(* IEC 61131-3 sources: daoli-st-library/DL_Motion (part 2) *)

(* ---- FB_DL_ResolverEncoderRedundSwitch.st ---- *)
(*
    FB_DL_ResolverEncoderRedundSwitch —— 旋变 + 增量编码器双通道角反馈冗余判定与无扰切换
    ------------------------------------------------------------------
    组件名    : FB_DL_ResolverEncoderRedundSwitch
    分类      : DL_Motion / Feedback Redundancy（反馈冗余切换）
    一句话功能: 双通道角反馈偏差超限时判定哪一路可信并无扰切到单通道运行，
                切换过程中输出角度受变率限制，绝不产生位置跳变。
    复杂度    : C4
    版本      : v1.0.0
    开源溯源  : 无（clean-room 自研，未借鉴任何开源实现）
    平台      : 纯 IEC 61131-3（TON / R_TRIG / ABS / REAL_TO_INT / INT_TO_REAL 标准转换），
                目标编译器 RuSTy 1.0.8，兼容 CODESYS 3.5 / TwinCAT 3 / 汇川 InoProShop /
                Machine Expert；无 PROPERTY、无 VLA、无 FOR..DOWNTO、无 AS 类方言
    ------------------------------------------------------------------
    功能说明  : ① 角差按 360° 环形折算：先各自折到 [0,360)，再
                   d := ABS(fAngleA − fAngleB)；IF d > 180 THEN d := 360 − d（结果域 [0,180]）；
                ② 双通道都有效且角差在容差内 → 融合输出（两路短弧中点），并每拍刷新
                   「融合参照角」_fRefDeg，供后续判定「哪一路可信」时作参照；
                ③ 角差超容差且持续 tFaultPersistMs（TON 无条件刷新）→ 判 SUSPECT；
                   任一路 bXValid = FALSE（或该路角度非有限）→ 直接判该路失效并切单通道；
                ④ 判定「哪一路可信」：以「最近一次双通道合格时的融合参照角」为准，
                   取与参照偏离较小者（相等时稳定优先取旋变 A）；无参照 → LOST，不猜；
                ⑤ 切换时 fAngleOut 按 fMaxSlewDegPerSec 限变率跟随目标角：环形带符号差值
                   先钳到 ±每拍步长再累加，故任何切换都不产生跳变；
                ⑥ 输出通道码 nActiveChannel：0 = 融合、1 = 旋变 A、2 = 编码器 B、-1 = 无。
    量纲链    : fAngleADeg [°] − fAngleBDeg [°] → 角差 [°]（经 360° 折算，域 [0,180]）；
                _fDevRatio = _fDevDeg [°] ÷ _fTolGuard [°] → 无因次 [-]（故与 1.0 直比判超限）；
                fMaxSlewDegPerSec [°/s] × DL_RE_SAMPLE_S [s] → 每拍最大角增量 [°]；
                _fDelta [°] 钳到 ±步长 [°] 后加到 _fOut [°] 再折回 [0,360) → fAngleOut [°]。
                全程无「角度与时间相加」「比例与角度相加」，量纲链逐段闭合。
    代理假设  : （R95 三句声明）① 代理值 = 常量 DL_RE_SAMPLE_S = 0.004 s，代表本 FB 所在
                任务的标称扫描周期；② 覆盖范围 = 2 ms ~ 10 ms 的周期任务（最坏 ±60% 误差只
                影响切换变率的平滑度，不改变安全判据的判定结果）；③ 覆盖不到的区间
                （< 1 ms 高速任务、事件任务、扫描周期抖动超 10 ms）由驱动层位置环限幅与伺服
                自身加速度限制负责，本件限变率只作二级防线。
    交付门槛  : 本件使用 REAL_TO_INT / INT_TO_REAL 标准转换做角度折圈，须在 CODESYS /
                TwinCAT / InoProShop 三平台各编译验证一次（R64）。
    状态机    : eInit(0) --双路有效且角差在容差内--> eDualOk(10)
                eInit --双路有效但角差超限--> eSuspect(20)；--仅一路有效--> eSingleA(30)/eSingleB(40)
                eDualOk --角差超容差持续 tFaultPersistMs 到（tonDev.Q）--> eSuspect
                eDualOk/eSuspect --A 失效--> eSingleB；--B 失效--> eSingleA
                eSuspect --有参照且可判--> eSingleA/eSingleB；--无参照或双路皆失效--> eLost(90)
                eSingleA/eSingleB --对侧恢复且一致计时到（tonAgree.Q）--> eDualOk
                eSingleA --A 失效--> eLost；eSingleB --B 失效--> eLost
                eLost --双路恢复且一致计时到（tonAgree.Q）--> eDualOk；
                eLost --单路恢复且确认计时到（tonSingle.Q）--> eSingleA/eSingleB（先进单通道，不直接回双通道）
                解除路径自证：tonSingle 的 IN 为「恰好一路可用」，故 eLost 的单路恢复边恒可达；
                若两路长期不一致且从未建立参照，eLost 按设计保持（不猜），bReset 重建参照后再裁决
    失能语义  : bEnable = FALSE 时 eState := eInit、nActiveChannel := -1、bLost := FALSE，
                fAngleOut 冻结保持末值（不跳变、不清零）；恢复使能后按变率追随新目标角。
                取「冻结保持」而非「降级清零」：角度是位置事实量，清零等于伪造位置（R191）。
    复位作用域: bReset 上升沿①清 _fRefDeg 与 _bRefValid（参照作废，须重建双通道合格）；
                ②清 _bCfgBad 与各成因位；③迁相回 eInit；④不清 _fOut（角度不得因复位跳变）。
    防御口径  : NaN 用自反 f<>f；±Inf 用 (f−f)<>(f−f)；另设幅值域闸 ABS(f) > 1.0E30。
                折圈除法的除子为常量 360.0（无零风险），但实数转整数前先做幅值域钳制，防
                REAL_TO_INT 溢出翻转（R151）；容差比值除法先以 DL_RE_TOL_FLOOR 两级兜底除子。
    规格补充  : 派单引脚表未含变率限制引脚，但设计要求「输出必须限变率」，故补充输入
                fMaxSlewDegPerSec（默认 3600 °/s，即 10 圈每秒）。派单写作 iActiveChannel（INT）；
                本库命名规范 1.2 规定有符号整数前缀为 n、i 专用于接口引用，故落为
                nActiveChannel，语义与码值一字不减。另按 R190 归因唯一补充 bCfgErr / bDataErr
                两个诊断位，使「组态非法」与「通道数据非有限」两条成因各自可观测。
    码位说明  : 本件按零码位范式交付，不分配 16# 事件码；失效成因（A 失效 / B 失效 /
                双路同时失效 / 无参照 / 当前通道失效 / 组态非法）各有独立内部成员，
                经 eState 与 bLost 观测，不共用同一枚举成员归因（R190）。
    修订记录  : 2026-11-24 v1.0.0 首次入库（R87 批 · #2）
*)
TYPE E_DL_ResEncState :
(
    eInit    := 0,    // 初始化或未投运：输出冻结，不判角差 | init or disabled, output frozen, no judging
    eDualOk  := 10,   // 双通道合格：融合输出，刷新融合参照角 | dual channels healthy, fused output, reference refreshed
    eSuspect := 20,   // 疑似：角差持续超容差，正在判定可信通道 | suspect, deviation persisted, arbitrating the trusted channel
    eSingleA := 30,   // 单通道 A：仅旋变通道参与输出 | single channel A, resolver only
    eSingleB := 40,   // 单通道 B：仅编码器通道参与输出 | single channel B, encoder only
    eLost    := 90    // 失效：无可信通道或无参照可判，输出冻结 | lost, no trusted channel or no reference
);
END_TYPE

FUNCTION_BLOCK FB_DL_ResolverEncoderRedundSwitch
VAR_INPUT
    bEnable            : BOOL;                    // 使能电平，TRUE = 允许切换判定 | enable level, TRUE = arbitration active
    bReset             : BOOL;                    // 复位请求，上升沿生效 | reset request, rising-edge active
    fAngleADeg         : REAL;                    // 旋变通道角度 [°]，任意圈数，内部折到 0..360 | resolver angle [deg]
    fAngleBDeg         : REAL;                    // 增量编码器角度 [°]，任意圈数，内部折到 0..360 | encoder angle [deg]
    fTolDeg            : REAL := 0.5;             // 双通道允许角差 [°]，须为正 | allowed channel deviation [deg]
    tFaultPersistMs    : TIME := T#100MS;         // 超限与恢复一致的持续确认时长 [ms] | persistence time [ms]
    bAValid            : BOOL;                    // 旋变通道有效位，驱动侧给出 | resolver channel validity from the drive
    bBValid            : BOOL;                    // 编码器通道有效位，驱动侧给出 | encoder channel validity from the drive
    fMaxSlewDegPerSec  : REAL := 3600.0;          // 输出角度最大变率 [°/s]，须为正 | max output slew rate [deg/s]
END_VAR
VAR_OUTPUT
    eState             : E_DL_ResEncState;        // 主状态，供 HMI 与联锁使用 | main state for HMI and interlocks
    fAngleOut          : REAL;                    // 参与位置环的输出角度 [°]，域 [0,360) 且限变率 | output angle [deg]
    fDeviationDeg      : REAL;                    // 本拍环形角差 [°]，域 [0,180] | circular deviation this scan [deg]
    nActiveChannel     : INT;                     // 通道码：0 融合 / 1 旋变 A / 2 编码器 B / -1 无 | channel code
    bSwitchEvent       : BOOL;                    // 通道切换事件位，单拍 | channel switch event, single scan
    bLost              : BOOL;                    // 失效汇总位，eLost 相为 TRUE | lost aggregate, TRUE in the eLost phase
    bCfgErr            : BOOL;                    // 组态非法诊断位（归因唯一，R190）| bad-configuration flag, unique attribution
    bDataErr           : BOOL;                    // 数据非有限诊断位（归因唯一，R190）| non-finite data flag, unique attribution
END_VAR
VAR
    rtReset            : R_TRIG;                  // 复位上升沿实例，每拍无条件刷新 | reset rising-edge instance
    tonDev             : TON;                     // 角差超限持续确认计时，每拍无条件刷新 | deviation persistence timer
    tonAgree           : TON;                     // 双通道一致确认计时，每拍无条件刷新 | agreement persistence timer
    tonSingle          : TON;                     // 单通道恢复确认计时，每拍无条件刷新 | single-channel recovery timer
    _eState            : E_DL_ResEncState := E_DL_ResEncState.eInit; // 状态机内部当前态 | internal current state
    _bInit             : BOOL := TRUE;            // 首扫初始化标志，含参照与输出保持槽状态 | first-scan init flag
    _bResetLatch       : BOOL := FALSE;           // 复位沿锁存量，本拍末清除 | reset-edge latch, cleared at scan end
    _bCfgBad           : BOOL := FALSE;           // 组态非法标志 | bad configuration flag
    _bAOk              : BOOL := FALSE;           // 旋变通道可用（有效位且角度有限）| resolver channel usable
    _bBOk              : BOOL := FALSE;           // 编码器通道可用（有效位且角度有限）| encoder channel usable
    _bLostBoth         : BOOL := FALSE;           // 双路同时失效成因位（归因唯一）| both channels lost
    _bNoRef            : BOOL := FALSE;           // 无融合参照成因位（归因唯一）| no reference available
    _bChLost           : BOOL := FALSE;           // 当前单通道失效成因位（归因唯一）| the active single channel was lost
    _fOut              : REAL := 0.0;             // 输出角度保持槽 [°]，域 [0,360) | output angle holder [deg]
    _fRefDeg           : REAL := 0.0;             // 融合参照角 [°]，仅在双通道合格时刷新 | fused reference angle [deg]
    _bRefValid         : BOOL := FALSE;           // 融合参照角可用标志 | fused reference valid flag
    _fDevDeg           : REAL := 0.0;             // 本拍环形角差 [°] | circular deviation this scan [deg]
    _fDevRatio         : REAL := 0.0;             // 角差与容差之比 [-]，判超限用 | deviation to tolerance ratio
    _fTolGuard         : REAL := 0.0;             // 带下限兜底的容差 [°]，作除法除子 | tolerance with floor, used as divisor
    _fSlewStep         : REAL := 0.0;             // 每拍最大角增量 [°] | max angle increment per scan [deg]
    _fDelta            : REAL := 0.0;             // 本拍待施加带符号角增量 [°]（已钳位）| clamped angle increment [deg]
    _fTarget           : REAL := 0.0;             // 本拍目标角 [°] | target angle this scan [deg]
    _fFuse             : REAL := 0.0;             // 本拍融合角 [°] | fused angle this scan [deg]
    _fDevA             : REAL := 0.0;             // A 相对参照的偏离 [°] | A deviation from the reference [deg]
    _fDevB             : REAL := 0.0;             // B 相对参照的偏离 [°] | B deviation from the reference [deg]
    _nCh               : INT := -1;               // 本拍通道码 | channel code this scan
    _nChPrev           : INT := -1;               // 上一拍通道码，供切换事件差分 | previous channel code for the switch event
    nFoldIdx           : INT := 0;                // 折圈方法内残余修正循环下标 | residue loop index inside the folding method
END_VAR
VAR CONSTANT
    DL_RE_EPS          : REAL := 1.0E-6;          // 浮点判零容差 [°] | float zero tolerance [deg]
    DL_RE_TOL_FLOOR    : REAL := 1.0E-4;          // 容差参数下限兜底 [°] | tolerance floor [deg]
    DL_RE_MAG_MAX      : REAL := 1.0E30;          // 有限幅值域闸上限（角度与变率）[°] | magnitude domain bound [deg]
    DL_RE_FOLD_MAX     : REAL := 1.0E6;           // 折圈前的角度幅值域上限 [°]，实数转整数前钳制 | fold domain bound [deg]
    DL_RE_SAMPLE_S     : REAL := 0.004;           // 代理扫描周期 [s]，见头注释代理假设三句 | proxy sample period [s]
    DL_RE_DEG_FULL     : REAL := 360.0;           // 整圈角度 [°] | full turn [deg]
    DL_RE_DEG_HALF     : REAL := 180.0;           // 半圈角度 [°] | half turn [deg]
    DL_RE_FUSE_W       : REAL := 0.5;             // 融合权重，两路等权且权值和为 1 [-] | fusion weight, sums to one
    DL_RE_CH_FUSE      : INT := 0;                // 通道码：融合 | channel code, fused
    DL_RE_CH_A         : INT := 1;                // 通道码：旋变 A | channel code, resolver A
    DL_RE_CH_B         : INT := 2;                // 通道码：编码器 B | channel code, encoder B
    DL_RE_CH_NONE      : INT := -1;               // 通道码：无 | channel code, none
    DL_RE_FOLD_ITER    : INT := 8;                // 折圈残余修正最大迭代次数（防死循环计数器）| fold iteration guard
END_VAR

METHOD FoldAngleDeg : REAL
(*
    角度折圈：把任意圈数角度折到 [0,360)。先按幅值域钳制再转整数，防 REAL_TO_INT 溢出翻转。
    Angle folding into [0,360): the magnitude is bounded before the real-to-integer conversion.
*)
VAR_INPUT
    fIn : REAL;                                   // 待折圈角度 [°] | angle to fold [deg]
END_VAR
VAR
    nTurn : INT;                                  // 整圈数，截断取整后按符号修正 [-] | whole turns after truncation
END_VAR
IF (fIn <> fIn) OR ((fIn - fIn) <> (fIn - fIn)) THEN
    FoldAngleDeg := 0.0;                          // NaN 或 ±Inf：返回哨兵零点，由调用方闸门拦截 | non-finite input returns the sentinel zero
    RETURN;
END_IF
IF (fIn > DL_RE_FOLD_MAX) OR (fIn < (0.0 - DL_RE_FOLD_MAX)) THEN
    FoldAngleDeg := 0.0;                          // 超折圈域：返回哨兵零点不猜，域外由上游闸门负责 | out of fold domain, return the sentinel
    RETURN;
END_IF
nTurn := REAL_TO_INT(fIn / DL_RE_DEG_FULL);       // 圈数 [-] = [°] ÷ 常量 360.0（除子为常量，无除零风险）| turns, constant divisor
FoldAngleDeg := fIn - INT_TO_REAL(nTurn) * DL_RE_DEG_FULL; // 折圈结果 [°] = [°] − [-] × [°] | folded angle [deg]
FOR nFoldIdx := 1 TO DL_RE_FOLD_ITER DO
    IF FoldAngleDeg < 0.0 THEN
        FoldAngleDeg := FoldAngleDeg + DL_RE_DEG_FULL; // 负角补整圈 [°] | add one turn for negative angles
    END_IF
END_FOR
IF FoldAngleDeg >= DL_RE_DEG_FULL THEN
    FoldAngleDeg := 0.0;                          // 折圈后仍越上界（数值极值退化）：返回哨兵零点 | degenerate result returns the sentinel
END_IF
END_METHOD

METHOD FoldDeviationDeg : REAL
(*
    环形角差幅值：d := ABS(A − B)；IF d > 180 THEN d := 360 − d，结果域 [0,180]（派单指定口径）。
    Circular deviation magnitude, exactly the formula requested by the dispatch.
*)
VAR_INPUT
    fAngleA : REAL;                               // A 通道角度 [°] | channel A angle [deg]
    fAngleB : REAL;                               // B 通道角度 [°] | channel B angle [deg]
END_VAR
VAR
    fD : REAL;                                    // 角差中间量 [°] | deviation intermediate [deg]
END_VAR
fD := ABS(FoldAngleDeg(fAngleA) - FoldAngleDeg(fAngleB)); // 折圈后作差取绝对值 [°] | absolute difference of folded angles
IF fD > DL_RE_DEG_HALF THEN
    fD := DL_RE_DEG_FULL - fD;                    // 折到短弧侧 [°]，与派单口径一致 | fold onto the short arc [deg]
END_IF
FoldDeviationDeg := fD;
END_METHOD

METHOD FoldSignedDiff : REAL
(*
    环形带符号差：返回 A − B 折到 (-180, 180]，用于融合与限变率增量计算。
    Signed circular difference folded into (-180, 180], used by fusion and by the slew limiter.
*)
VAR_INPUT
    fAngleA : REAL;                               // 被减角度 [°] | minuend angle [deg]
    fAngleB : REAL;                               // 减数角度 [°] | subtrahend angle [deg]
END_VAR
VAR
    fD : REAL;                                    // 带符号角差中间量 [°] | signed difference intermediate [deg]
END_VAR
fD := FoldAngleDeg(fAngleA) - FoldAngleDeg(fAngleB); // 折圈后作差 [°] | difference of folded angles [deg]
IF fD > DL_RE_DEG_HALF THEN
    fD := fD - DL_RE_DEG_FULL;                    // 折到负侧 [°] | fold into the negative side [deg]
END_IF
IF fD <= (0.0 - DL_RE_DEG_HALF) THEN
    fD := fD + DL_RE_DEG_FULL;                    // 折到正侧 [°] | fold into the positive side [deg]
END_IF
FoldSignedDiff := fD;
END_METHOD

// 段 1｜输出安全侧预置与首扫初始化（含参照与保持槽状态，故必须有 _bInit，R310）
// segment 1, safe-value presets and first-scan initialisation; the reference holder requires _bInit
nActiveChannel := DL_RE_CH_NONE;                   // 预置通道码「无」| preset channel code to none
bLost := FALSE;                                    // 预置未失效 | preset not lost
bSwitchEvent := FALSE;                             // 预置无切换事件 | preset no switch event
_fDevDeg := 0.0;                                   // 预置角差 0 [°] | preset zero deviation [deg]
_fDevRatio := 0.0;                                 // 预置角差比 0 [-] | preset zero ratio
_bCfgBad := FALSE;                                 // 预置组态合法 | preset legal configuration
_bLostBoth := FALSE;                               // 预置双路未同时失效 | preset both channels not lost
_bNoRef := FALSE;                                  // 预置参照缺失未置位 | preset reference-missing flag clear
_bChLost := FALSE;                                 // 预置当前通道未失效 | preset active-channel-lost flag clear
_nCh := DL_RE_CH_NONE;                             // 预置本拍通道码「无」| preset the channel code to none
IF _bInit THEN
    _bInit := FALSE;                               // 首扫只执行一次 | runs once on the first scan
    _eState := E_DL_ResEncState.eInit;             // 首扫状态回初相 | initialise the state
    _bRefValid := FALSE;                           // 参照角作废，须重建 | invalidate the reference
    IF (fAngleADeg <> fAngleADeg) OR ((fAngleADeg - fAngleADeg) <> (fAngleADeg - fAngleADeg)) THEN
        _fOut := 0.0;                              // 首扫角度非有限：保持槽取哨兵零点，等闸门置失效 | non-finite first angle
    ELSE
        _fOut := FoldAngleDeg(fAngleADeg);         // 首扫以旋变角为输出起点 [°]，避免首拍从 0 跳变 | start from the resolver angle
    END_IF
    _nChPrev := DL_RE_CH_NONE;                     // 首扫通道快照为「无」| first-scan channel snapshot
END_IF

// 段 2｜通道可用性判定：有效位 + NaN 自反 + Inf 自减 + 幅值域，逐个浮点入参枚举（R4 / R151 / R272）
// segment 2, channel usability: validity bit plus NaN self-reflexive, Inf self-subtraction and the magnitude bound
_bAOk := bAValid;
IF (fAngleADeg <> fAngleADeg) OR ((fAngleADeg - fAngleADeg) <> (fAngleADeg - fAngleADeg)) THEN
    _bAOk := FALSE;                                // 旋变角 NaN 或 ±Inf：判该路失效 | NaN or infinity, the channel is unusable
END_IF
IF ABS(fAngleADeg) > DL_RE_MAG_MAX THEN
    _bAOk := FALSE;                                // 旋变角超幅值域：判该路失效 | beyond the magnitude domain, unusable
END_IF
_bBOk := bBValid;
IF (fAngleBDeg <> fAngleBDeg) OR ((fAngleBDeg - fAngleBDeg) <> (fAngleBDeg - fAngleBDeg)) THEN
    _bBOk := FALSE;                                // 编码器角 NaN 或 ±Inf：判该路失效 | NaN or infinity, the channel is unusable
END_IF
IF ABS(fAngleBDeg) > DL_RE_MAG_MAX THEN
    _bBOk := FALSE;                                // 编码器角超幅值域：判该路失效 | beyond the magnitude domain, unusable
END_IF

// 段 3｜容差两级兜底与组态闸（容差作除子，必须先兜底再除；变率须为正且有限）
// segment 3, two-stage tolerance fallback and configuration gate; the tolerance is a divisor, floor it first
_fTolGuard := fTolDeg;                             // 取配置容差 [°] | take the configured tolerance [deg]
IF (fTolDeg <> fTolDeg) OR ((fTolDeg - fTolDeg) <> (fTolDeg - fTolDeg)) THEN
    _fTolGuard := DL_RE_TOL_FLOOR;                 // 容差非有限：一级回默认下限 [°] | non-finite tolerance falls back to the floor
END_IF
IF _fTolGuard < DL_RE_TOL_FLOOR THEN
    _fTolGuard := DL_RE_TOL_FLOOR;                 // 容差过小或为负：二级按有效域钳定 [°] | too small or negative, clamp to the floor
END_IF
IF (fMaxSlewDegPerSec <> fMaxSlewDegPerSec) OR ((fMaxSlewDegPerSec - fMaxSlewDegPerSec) <> (fMaxSlewDegPerSec - fMaxSlewDegPerSec)) THEN
    _bCfgBad := TRUE;                              // 变率非有限：组态非法 | non-finite slew rate, illegal configuration
END_IF
IF fMaxSlewDegPerSec <= DL_RE_EPS THEN
    _bCfgBad := TRUE;                              // 变率非正：组态非法（无变率限制即失去无扰切换保障）| non-positive slew rate
END_IF
IF ABS(fMaxSlewDegPerSec) > DL_RE_MAG_MAX THEN
    _bCfgBad := TRUE;                              // 变率超幅值域：组态非法 | slew rate beyond the magnitude domain
END_IF
IF tFaultPersistMs < T#0S THEN
    _bCfgBad := TRUE;                              // 持续确认时长为负：组态非法 | negative persistence time, illegal configuration
END_IF

// 段 4｜本拍角差与角差比（双路都可用才计算，否则记 0 且不参与判据）
// segment 4, deviation and deviation ratio this scan; computed only when both channels are usable
IF _bAOk AND _bBOk THEN
    _fDevDeg := FoldDeviationDeg(fAngleADeg, fAngleBDeg); // 环形角差 [°] | circular deviation [deg]
    _fDevRatio := _fDevDeg / _fTolGuard;           // 角差比 [-] = [°] ÷ [°]，_fTolGuard 已两级兜底非零 | guarded division
ELSE
    _fDevDeg := 0.0;                               // 单路或双路失效：角差无意义记 0 [°] | deviation meaningless here
    _fDevRatio := 0.0;                             // 单路或双路失效：角差比记 0 [-] | ratio meaningless here
END_IF

// 段 5｜定时器与沿实例无条件周期刷新（R7：严禁放入 IF / CASE 分支内部），入参为本拍已算量
// segment 5, timers and edge instances refreshed unconditionally, fed with values already computed this scan
rtReset(CLK := bReset);
tonDev(IN := bEnable AND _bAOk AND _bBOk AND (_fDevRatio > 1.0), PT := tFaultPersistMs);
tonAgree(IN := bEnable AND _bAOk AND _bBOk AND (_fDevRatio <= 1.0), PT := tFaultPersistMs);
tonSingle(IN := bEnable AND (_bAOk OR _bBOk) AND (NOT (_bAOk AND _bBOk)), PT := tFaultPersistMs);
IF rtReset.Q THEN
    _bResetLatch := TRUE;                          // 复位沿存锁存量，段 6 统一消费 | store the reset edge, consumed in segment 6
END_IF

// 段 6｜复位沿处理（先复位后判据，保证本拍新事件不被抹除，R275）
// segment 6, reset edge handling; reset runs before the criteria so same-scan events survive
IF _bResetLatch THEN
    _bRefValid := FALSE;                           // 参照作废，须重新建立双通道合格 | invalidate the reference
    _fRefDeg := 0.0;                               // 参照角清零 [°] | clear the reference angle [deg]
    _bCfgBad := FALSE;                             // 清组态非法标志（下一拍按新参数重判）| clear the configuration flag
    _eState := E_DL_ResEncState.eInit;             // 迁回初相 | return to the init phase
    _nCh := DL_RE_CH_NONE;                         // 复位拍通道码置无 | channel code set to none on the reset scan
END_IF

// 段 7｜组态非法：无变率限制即无法保证无扰切换，组态闸优先于一切判定
// segment 7, illegal configuration: without a slew limit the bumpless switch cannot be guaranteed
IF _bCfgBad THEN
    _eState := E_DL_ResEncState.eLost;
END_IF

// 段 8｜主状态机：ENUM + CASE + ELSE 兜底（R6）
// segment 8, main state machine with ENUM + CASE + ELSE fallback
CASE _eState OF
E_DL_ResEncState.eInit:
    _fTarget := _fOut;                             // 初相不追随目标，输出冻结 [°] | the init phase does not chase a target
    // 拍 N 进入：首扫、复位沿或使能撤除；本拍行为：只做有效性分类，不改输出角；
    // 拍 N+1 转出：双路有效且角差在容差内 → eDualOk；双路有效但超容差 → eSuspect；
    //              仅一路有效 → eSingleA / eSingleB；两路皆失效 → eLost
    // entered on the first scan, the reset edge or on disable; only classifies validity and never moves the output;
    // exits to eDualOk, eSuspect, eSingleA, eSingleB or eLost according to the validation result
    IF bEnable THEN
        IF _bAOk AND _bBOk THEN
            IF _fDevRatio <= 1.0 THEN
                _eState := E_DL_ResEncState.eDualOk;
            ELSE
                _eState := E_DL_ResEncState.eSuspect;
            END_IF
        ELSIF _bAOk THEN
            _eState := E_DL_ResEncState.eSingleA;
        ELSIF _bBOk THEN
            _eState := E_DL_ResEncState.eSingleB;
        ELSE
            _bLostBoth := TRUE;                    // 双路同时失效（独立成因）| both channels lost, unique attribution
            _eState := E_DL_ResEncState.eLost;
        END_IF
    END_IF

E_DL_ResEncState.eDualOk:
    // 融合：以 A 为基准加半幅带符号差，权重和为 1，故结果恒落在两路短弧中点
    // fusion: start from A and add half of the signed difference, giving the short-arc midpoint
    _fFuse := FoldAngleDeg(fAngleADeg + FoldSignedDiff(fAngleBDeg, fAngleADeg) * DL_RE_FUSE_W); // 融合角 [°] | fused angle [deg]
    _fTarget := _fFuse;                            // 双通道相目标为融合角 [°] | target is the fused angle
    _nCh := DL_RE_CH_FUSE;                         // 通道码：融合 | channel code fused
    _fRefDeg := _fFuse;                            // 刷新融合参照角 [°]，供后续判可信通道 | refresh the fused reference [deg]
    _bRefValid := TRUE;                            // 参照角已建立 | reference established
    IF NOT bEnable THEN
        _eState := E_DL_ResEncState.eInit;          // 失能回初相（输出冻结）| disable returns to init
    ELSIF (NOT _bAOk) AND (NOT _bBOk) THEN
        _bLostBoth := TRUE;                        // 双路同时失效 | both channels lost
        _eState := E_DL_ResEncState.eLost;
    ELSIF NOT _bAOk THEN
        _eState := E_DL_ResEncState.eSingleB;       // 旋变失效 → 切编码器 | resolver lost, switch to the encoder
    ELSIF NOT _bBOk THEN
        _eState := E_DL_ResEncState.eSingleA;       // 编码器失效 → 切旋变 | encoder lost, switch to the resolver
    ELSIF tonDev.Q THEN
        _eState := E_DL_ResEncState.eSuspect;       // 角差超容差持续确认到 → 进疑似相 | persisted deviation, enter suspect
    END_IF

E_DL_ResEncState.eSuspect:
    _fTarget := _fOut;                             // 疑似相不追随任何通道，输出冻结等裁决 [°] | no channel is chased here
    _nCh := DL_RE_CH_NONE;                         // 疑似相无有效通道码 | no valid channel code in suspect
    IF NOT bEnable THEN
        _eState := E_DL_ResEncState.eInit;          // 失能回初相 | disable returns to init
    ELSIF _bAOk AND _bBOk THEN
        IF _fDevRatio <= 1.0 THEN
            _eState := E_DL_ResEncState.eDualOk;   // 角差已回到容差内：撤销疑似，无需切换 | deviation back inside, cancel the suspect
        ELSIF _bRefValid THEN
            _fDevA := FoldDeviationDeg(fAngleADeg, _fRefDeg); // A 相对参照偏离 [°] | A deviation from the reference [deg]
            _fDevB := FoldDeviationDeg(fAngleBDeg, _fRefDeg); // B 相对参照偏离 [°] | B deviation from the reference [deg]
            IF (_fDevA < _fDevB) OR (_fDevA = _fDevB) THEN
                _eState := E_DL_ResEncState.eSingleA; // 取偏离小者；相等时稳定优先保留旋变 A | closer channel wins, ties keep the resolver
            ELSE
                _eState := E_DL_ResEncState.eSingleB;
            END_IF
        ELSE
            _bNoRef := TRUE;                       // 无参照可判：不猜（独立成因）| no reference, refuse to guess
            _eState := E_DL_ResEncState.eLost;
        END_IF
    ELSIF _bAOk THEN
        _eState := E_DL_ResEncState.eSingleA;       // 仅旋变可用 | only the resolver is usable
    ELSIF _bBOk THEN
        _eState := E_DL_ResEncState.eSingleB;       // 仅编码器可用 | only the encoder is usable
    ELSE
        _bLostBoth := TRUE;                        // 双路同时失效 | both channels lost
        _eState := E_DL_ResEncState.eLost;
    END_IF

E_DL_ResEncState.eSingleA:
    _fTarget := FoldAngleDeg(fAngleADeg);          // 单通道 A：目标为旋变角 [°] | single A, target is the resolver angle
    _nCh := DL_RE_CH_A;                            // 通道码：旋变 A | channel code A
    IF NOT bEnable THEN
        _eState := E_DL_ResEncState.eInit;          // 失能回初相 | disable returns to init
    ELSIF NOT _bAOk THEN
        _bChLost := TRUE;                          // 当前通道失效（独立成因）：不切换、直接失效 | the active channel is lost
        _eState := E_DL_ResEncState.eLost;
    ELSIF _bBOk AND tonAgree.Q THEN
        _eState := E_DL_ResEncState.eDualOk;        // 对侧恢复且一致计时到 → 回双通道 | peer recovered and agreed, back to dual
    END_IF

E_DL_ResEncState.eSingleB:
    _fTarget := FoldAngleDeg(fAngleBDeg);          // 单通道 B：目标为编码器角 [°] | single B, target is the encoder angle
    _nCh := DL_RE_CH_B;                            // 通道码：编码器 B | channel code B
    IF NOT bEnable THEN
        _eState := E_DL_ResEncState.eInit;          // 失能回初相 | disable returns to init
    ELSIF NOT _bBOk THEN
        _bChLost := TRUE;                          // 当前通道失效（独立成因）：不切换、直接失效 | the active channel is lost
        _eState := E_DL_ResEncState.eLost;
    ELSIF _bAOk AND tonAgree.Q THEN
        _eState := E_DL_ResEncState.eDualOk;        // 对侧恢复且一致计时到 → 回双通道 | peer recovered and agreed, back to dual
    END_IF

E_DL_ResEncState.eLost:
    _fTarget := _fOut;                             // 失效相冻结输出，宁可保持也不跳变 [°] | frozen output, never jump
    _nCh := DL_RE_CH_NONE;                         // 无有效通道码 | no valid channel code
    IF NOT bEnable THEN
        _eState := E_DL_ResEncState.eInit;          // 失能回初相 | disable returns to init
    ELSIF _bAOk AND _bBOk AND tonAgree.Q THEN
        _eState := E_DL_ResEncState.eDualOk;        // 双路恢复且一致计时到 → 回双通道 | both recovered and agreed
    ELSIF _bAOk AND tonSingle.Q THEN
        _eState := E_DL_ResEncState.eSingleA;       // 单路 A 恢复且确认到 → 先切单通道（不直接回双通道）| single A confirmed
    ELSIF _bBOk AND tonSingle.Q THEN
        _eState := E_DL_ResEncState.eSingleB;       // 单路 B 恢复且确认到 → 先切单通道 | single B confirmed
    END_IF
    // 解除路径自证：tonSingle 的 IN = 恰好一路可用，故上式在「单路恢复」场景恒可达；
    // 若两路长期不一致且无参照，本相按设计保持（不猜），bReset 可重建参照后重新裁决。

ELSE
    // 非法枚举值（越界或未定义成员）：不猜，冻结输出并置失效相
    // illegal enumerator: no guessing, freeze the output and fall into the lost phase
    _fTarget := _fOut;
    _nCh := DL_RE_CH_NONE;
    _eState := E_DL_ResEncState.eLost;
END_CASE;

// 段 9｜限变率追随：环形带符号差先钳到 ±每拍步长再累加，故任何切换都不产生跳变
// segment 9, slew-limited tracking; the circular difference is clamped to the per-scan step before integration
IF bEnable AND (NOT _bCfgBad) THEN
    _fSlewStep := fMaxSlewDegPerSec * DL_RE_SAMPLE_S; // 每拍最大角增量 [°] = [°/s] × [s] | per-scan step [deg]
    _fDelta := FoldSignedDiff(_fTarget, _fOut);    // 待施加带符号角增量 [°] | signed increment to apply [deg]
    IF _fDelta > _fSlewStep THEN
        _fDelta := _fSlewStep;                     // 正向钳到步长上限 [°] | clamp to the positive step
    END_IF
    IF _fDelta < (0.0 - _fSlewStep) THEN
        _fDelta := 0.0 - _fSlewStep;               // 负向钳到步长下限 [°] | clamp to the negative step
    END_IF
    _fOut := FoldAngleDeg(_fOut + _fDelta);        // 累加并折圈 [°] | integrate and fold [deg]
END_IF
// 失能或组态非法时 _fOut 冻结保持末值（头注释已声明「冻结保持」语义，R191）

// 段 10｜出口单点映射（切换事件由通道码差分派生，单拍；快照在本段末更新）
// segment 10, single-point output mapping; the switch event is derived from the channel code difference
eState := _eState;                                 // 状态映射 | state mapping
fAngleOut := _fOut;                                // 输出角度映射 [°] | output angle mapping [deg]
fDeviationDeg := _fDevDeg;                         // 角差映射 [°] | deviation mapping [deg]
nActiveChannel := _nCh;                            // 通道码映射 | channel code mapping
bSwitchEvent := (_nCh <> _nChPrev);                // 切换单拍位 = 本拍码与上拍码不同 | one-scan switch pulse
_nChPrev := _nCh;                                  // 更新通道码快照（非清零，仅供下一拍差分）| update the snapshot
bLost := (_eState = E_DL_ResEncState.eLost);       // 失效汇总由状态派生 | lost aggregate derived from the state
bCfgErr := _bCfgBad;                               // 组态非法诊断位 | bad-configuration diagnostic
bDataErr := (NOT _bAOk) OR (NOT _bBOk);            // 数据非有限诊断位（通道可用性直接派生）| non-finite data diagnostic

// 段 11｜本拍消费量收尾（仅清沿锁存；不触碰任何锁存位与 CASE 内写入量）
// segment 11, end-of-scan cleanup; only the edge latch is cleared
_bResetLatch := FALSE;
END_FUNCTION_BLOCK

(* ---- FB_DL_VirtualMasterAxis.st ---- *)
(*
    FB_DL_VirtualMasterAxis —— 虚拟主轴相位源
    ------------------------------------------------------------------
    分类      : DL_Motion / MasterSource
    前缀      : FB_DL_
    版本      : 1.0.1
    溯源      : T2-4 S7 Motion 工艺对象分型（只借「同步轴需要独立主值源」的公开架构语义）；
                T1-6 PLCopen 凸轮/齿轮需要连续相位主值的公开条款为次源；
                斜坡积分器、精度门限、冻结策略与码位 100% 自有；clean-room 重写，
                未复制任何闭源厂商源码，参考实现仅限 MIT/Apache 许可
    道莅 clean-room 防御性实现：语义借鉴、代码与码位 100% 自有
    平台      : 纯 IEC 61131-3，CODESYS V3.5+ / TwinCAT 3 / InoProShop / Machine Expert 通用
    作者      : 道莅代码库 · PLC编程专家（R22 批 4 · #13）
    ------------------------------------------------------------------
    功能说明  : 电子凸轮 / 电子齿轮的主值源：把「速度给定 + 加减速限值」积分成连续相位、
                速度与加速度三个量，供从轴按相位跟随。本件不发任何运动指令、
                不自造轴状态枚举——它只回答「主轴现在在哪、多快、加速度多大」。
    相位精度  : 相位以 LREAL 累加。IEEE 754 双精度在 |x| > 1.0E15 mm 时相邻可表示
                差值已大于 1e-3 mm 量级，凸轮相位已失真而调用方看不出来，因此本件把
                1.0E15 设为硬门限：越限即报故障 02EE 并冻结相位，不静默累计。
                冻结而不是清零，是为了让调用方看清「停在哪」再决定复位。
    两条律    : ① bHold 走减速斜坡降到 0，绝不瞬时归零（瞬时归零会让从轴指令跳变）；
                ② 失能（bEnable 落）同样走减速斜坡，且残速期间相位继续积分，
                   因为轴物理上仍在走，位置不跟着走就等于伪造相位。
    设计取舍  : 复位沿优先于失能判定——同一拍既给 bPhaseReset 又撤 bEnable 时先复位再判状态，
                否则复位沿会被失能分支吞掉，调用方会以为「按了没反应」。
                参数类与非有限类故障（02ED）一律冻结速度与相位，不做「按末次速度继续跑」：
                采样周期不可信时继续积分等于用错误的 dt 编造相位。
    职责边界  : 本件只做「主值源」。主轴的使能、抱闸、限位、回零仍归轴功能块；
                本件不消费、不改写任何轴状态；Blending 速度融合不在本件能力范围。
    错误码    : 16#0004_01D7 加速度限幅生效（仍在斜坡中，未达给定）——信息级，边沿发布
                16#0004_01D8 相位复位已执行——信息级，单拍发布
                16#0004_02ED 采样周期非正 / 速度与限值参数非法或非有限——故障级，
                             冻结速度与相位并保持末次有效速度
                16#0004_02EE 相位累计超 LREAL 有效精度 1.0E15 mm，已冻结——故障级，
                             需调用方给 bPhaseReset 复位后才允许回待机
                16#0004_02EF 状态机落 ELSE 兜底（非法状态）——故障级，回 eFault
    码位总账  : 16#0004_01D7 用 / 16#0004_01D8 用 ｜ 16#0004_02ED 用 / 16#0004_02EE 用 / 16#0004_02EF 用
    状态机    : E_DL_VMasterState（eIdle / eRamping / eSteady / eHolding / eFault），
                CASE 含 ELSE 兜底，ELSE 置 16#0004_02EF 并回 eFault；
                斜坡与积分在本体段 6 执行，故障拍与故障相（eFault）均冻结，
                参数修复后须经失能复位或 bPhaseReset 才恢复积分（v1.0.1 终审修复）。
    采样约定  : fbPhaseReset 在本体首部无条件刷新（R40）；dt 由 tSample 引脚换算，
                严禁读取系统时钟；换算链 TIME_TO_DINT → DINT_TO_REAL 在
                CODESYS V3.5 / TwinCAT 3 / InoProShop / Machine Expert 四平台均为
                标准运算符，若目标平台仅实现 TIME_TO_REAL 可等价替换（编译门槛已声明）。
    依赖      : 仅 Standard.library（R_TRIG / LIMIT / ABS），不引用任何其他 DL_ 子库。
    验收向量  :
                V1 域外早退：tSample = T#0MS → 02ED、bError=TRUE、bValid=FALSE，
                   相位与速度两拍完全相同（冻结）。
                V2 上限限幅：fVelSet = 5000 mm/s、fAccLimit = 1000 mm/s²、tSample = 1 ms
                   → 每拍速度增量恰为 1.0 mm/s、bLimited=TRUE、01D7 只出现一拍。
                V3 跨段时序：eSteady 中 bHold 置位 → 速度按 fDecLimit 逐拍递减，
                   位置继续积分直到速度为 0 才停；不得出现速度阶跃为 0。
                V4 复位首拍：bPhaseReset 与撤 bEnable 同拍 → 复位优先执行
                   （fMasterPos = fPosInit、fMasterVel = 0、01D8），随后才回 eIdle。
    红线自检  : 1 全局变量声明零使用 / 外部变量访问零使用 / 物理地址零使用 —— 通过，全部量经引脚注入
                2 纯 IEC 61131-3 跨平台 —— 通过，仅 Standard.library，换算链已在头注释声明门槛
                3 防御性编程 —— 通过，浮点判等用 1.0E-6 容差、除法前判 dt > 0、无非有限穿透
                4 声明行同行中英双语注释 + 单位 —— 通过，逐行附注（含枚举成员）
                5 ENUM + CASE 且含 ELSE 兜底 —— 通过
                6 TON / R_TRIG 无条件刷新 —— 通过，段 1 先行调用
                7 无魔法数 —— 通过，门限与容差全部 VAR CONSTANT，时间为引脚
    修订记录  : 2026-11-16 v1.0.0 首次入库（R22 批 4 · #13）
                2026-11-16 v1.0.1 R22 终审修复：段 6 积分增加 eFault 相位门控——
                原实现中 eFault 态下 bError 仅在故障检出拍为真，参数修复后下一拍
                bError 归假即恢复积分，与「eFault 冻结速度与相位」的头注释承诺矛盾；
                修复后故障相彻底冻结，恢复仅经「失能复位」或「bPhaseReset」两条路径
*)
TYPE E_DL_VMasterState :
(
    eIdle    := 0,       // 未使能；若仍有残速则按减速限值降到零并继续积分 / not enabled, a residual velocity is ramped down and the phase keeps integrating
    eRamping := 10,      // 斜坡中，速度尚未达到给定 / ramping, the velocity has not reached the setpoint yet
    eSteady  := 20,      // 已达给定，速度稳定，bReady 置位 / at the setpoint, bReady is asserted
    eHolding := 30,      // 保持相，目标速度强制为 0 但按减速斜坡逼近 / holding, the target is forced to zero and approached through the deceleration ramp
    eFault   := 40       // 故障，速度与相位冻结 / fault, both velocity and phase are frozen
);
END_TYPE

FUNCTION_BLOCK FB_DL_VirtualMasterAxis
VAR_INPUT
    bEnable      : BOOL;                       // 使能，FALSE 时目标速度归零并走减速斜坡 / enable, FALSE forces the target to zero through the deceleration ramp
    fVelSet      : REAL;                       // 主轴速度给定 [mm/s]，非有限即拒绝 / master velocity setpoint [mm/s], a non-finite value is rejected
    fAccLimit    : REAL := 1000.0;             // 加速限值 [mm/s²]，必须大于 0 / acceleration limit [mm/s²], must exceed zero
    fDecLimit    : REAL := 1000.0;             // 减速限值 [mm/s²]，必须大于 0 / deceleration limit [mm/s²], must exceed zero
    bHold        : BOOL;                       // 保持，TRUE 时按减速斜坡降到 0 而非瞬时归零 / hold, TRUE ramps the velocity down instead of stepping it to zero
    bPhaseReset  : BOOL;                       // 相位复位，上升沿生效且优先于失能判定 / phase reset, effective on the rising edge and prior to the disable test
    fPosInit     : REAL := 0.0;                // 复位目标相位 [mm]，非有限即拒绝 / reset target phase [mm], a non-finite value is rejected
    tSample      : TIME := T#1MS;              // 采样周期 [ms]，必须大于 0，禁读系统时钟 / sample period [ms], must exceed zero, never read from the system clock
END_VAR
VAR_OUTPUT
    fMasterPos   : LREAL;                      // 主轴相位 [mm]，LREAL 累加 / master phase [mm], accumulated in LREAL
    fMasterVel   : REAL;                       // 主轴速度 [mm/s]，斜坡输出 / master velocity [mm/s], the ramp output
    fMasterAcc   : REAL;                       // 主轴加速度 [mm/s²]，本拍实际生效值 / master acceleration [mm/s²], the value actually applied this scan
    bReady       : BOOL;                       // 主值可用，速度已达给定（或保持相已停稳）/ master value usable, the velocity has reached the setpoint or the hold has settled
    bLimited     : BOOL;                       // 本拍被加减速限值截断 / this scan was clipped by an acceleration or deceleration limit
    eErr         : UDINT;                      // 错误码，0 表示无错 / error code, 0 means no error
    bError       : BOOL;                       // 故障级标志，仅故障级错误置位 / fault-class flag, set only on fault-level codes
    bValid       : BOOL;                       // 输出可用标志，= NOT bError / outputs valid flag, equals NOT bError
END_VAR
VAR
    fbPhaseReset  : R_TRIG;                    // 复位沿检测实例，本体首部无条件刷新 / reset edge instance, refreshed unconditionally
    _fPosL        : LREAL;                     // 相位累加器（本件唯一的跨周期状态）/ the phase accumulator, the only truly cyclic state of this block
    _fVel         : REAL;                      // 速度状态，斜坡积分结果 [mm/s] / velocity state, the ramp integration result [mm/s]
    _fTarget      : REAL;                      // 本拍有效目标速度（含失能与保持折算）[mm/s] / effective target velocity of this scan including disable and hold [mm/s]
    _fDtSec       : REAL;                      // 本拍采样周期折算秒值 [s] / sample period converted to seconds [s]
    _fMaxUp       : REAL;                      // 本拍允许的速度上升量 [mm/s] / permitted velocity increase of this scan [mm/s]
    _fMaxDn       : REAL;                      // 本拍允许的速度下降量 [mm/s] / permitted velocity decrease of this scan [mm/s]
    _fDiff        : REAL;                      // 目标与当前速度之差 [mm/s] / difference between the target and the current velocity [mm/s]
    _fDelta       : REAL;                      // 本拍速度增量，限幅后 [mm/s] / velocity increment of this scan after clipping [mm/s]
    _bParamBad    : BOOL;                      // 参数或采样非法标志 / illegal parameter or sample flag
    _bLimitPrev   : BOOL;                      // 上一拍限幅标志，用于信息码边沿发布 / previous-scan limiting flag used for the edge-published info code
    _eState       : E_DL_VMasterState;         // 当前状态 / current state
END_VAR
VAR CONSTANT
    DL_VM_MS_PER_S    : REAL := 1000.0;        // 毫秒与秒的换算系数 [ms/s] / milliseconds per second [ms/s]
    DL_VM_POS_MAX     : LREAL := 1.0E15;       // 相位有效精度上限 [mm]，越限即冻结 / effective phase precision limit [mm], exceeded means freeze
    DL_VM_INF_GUARD   : REAL := 4.0E38;        // REAL 非有限幅值判定阈（大于 REAL 最大值）[mm/s] / REAL non-finite magnitude guard [mm/s]
    DL_VM_EPS         : REAL := 1.0E-6;        // 速度判等容差 [mm/s] / velocity equality tolerance [mm/s]
    DL_VM_ZERO        : REAL := 0.0;           // 零值常量，避免裸字面量 [无量纲] / zero constant, avoids a bare literal [dimensionless]
    DL_VM_T_ZERO      : TIME := T#0S;          // 零时间常量，用于采样周期门禁 / zero time constant used by the sample gate
END_VAR

// 段 1｜复位沿实例无条件周期刷新（红线 6：严禁放入 IF / CASE）/ segment 1, unconditional edge refresh
fbPhaseReset(CLK := bPhaseReset);

// 段 2｜输出与错误状态预置 / segment 2, preset outputs and error status
eErr := 0;                                      // 预置无错误 / preset no error
bError := FALSE;                                // 预置无故障标志 / preset no error flag
bLimited := FALSE;                              // 预置本拍无限幅 / preset no limiting this scan
bReady := FALSE;                                // 预置主值不可用 / preset the master value as not usable
fMasterAcc := DL_VM_ZERO;                       // 预置本拍加速度为 0 / preset the applied acceleration to zero

// 段 3｜参数与采样门禁：① 采样周期非正 ② 限值非正或非有限 ③ 给定与复位值非有限
// segment 3, parameter and sample gate
_bParamBad := FALSE;                            // 先假定参数合法 / assume legal parameters first
IF (tSample <= DL_VM_T_ZERO)
   OR (fAccLimit <= DL_VM_ZERO)
   OR (fDecLimit <= DL_VM_ZERO) THEN
    _bParamBad := TRUE;                         // 采样周期或限值非正 / the sample period or a limit is not positive
END_IF

// 非有限检测：NaN 用自不自等捕获，±Inf 用幅值门捕获（REAL 最大约 3.4E38）
// non-finite detection, NaN via self-inequality and plus/minus infinity via the magnitude guard
IF (fVelSet - fVelSet) <> (fVelSet - fVelSet) THEN
    _bParamBad := TRUE;                         // 速度给定为 NaN / the velocity setpoint is NaN
ELSIF ABS(fVelSet) > DL_VM_INF_GUARD THEN
    _bParamBad := TRUE;                         // 速度给定为 ±Inf / the velocity setpoint is infinite
END_IF
IF (fPosInit - fPosInit) <> (fPosInit - fPosInit) THEN
    _bParamBad := TRUE;                         // 复位相位为 NaN / the reset phase is NaN
ELSIF ABS(fPosInit) > DL_VM_INF_GUARD THEN
    _bParamBad := TRUE;                         // 复位相位为 ±Inf / the reset phase is infinite
END_IF

IF _bParamBad THEN
    eErr := 16#0004_02ED;                       // 故障级：采样周期或速度参数非法 / fault: sample period or velocity parameter illegal
    bError := TRUE;                             // 置故障标志 / raise the fault flag
    _eState := E_DL_VMasterState.eFault;        // 转故障，本拍不积分 / go to fault, no integration this scan
    fMasterVel := _fVel;                        // 保持末次有效速度 [mm/s] / hold the last valid velocity [mm/s]
    bValid := FALSE;                            // 输出不可用 / outputs are not valid
END_IF

// 段 4｜有效目标速度：失能或保持都折算为 0，由斜坡逼近而非阶跃
// segment 4, effective target velocity; disable and hold both map to zero and are approached through the ramp
IF (NOT bEnable) OR bHold OR bError THEN
    _fTarget := DL_VM_ZERO;                     // 失能 / 保持 / 故障：目标为 0 / disabled, holding or faulted, the target is zero
ELSE
    _fTarget := fVelSet;                        // 正常运行：目标即给定 / normal operation, the target is the setpoint
END_IF

// 段 5｜相位复位：优先于失能判定（同一拍两者同时到达时先复位，否则沿被吞掉）
// segment 5, phase reset evaluated before the disable test so a joint edge is never swallowed
IF fbPhaseReset.Q AND (NOT _bParamBad) THEN
    _fPosL := fPosInit;                         // 相位直接置到复位目标 / the phase jumps to the reset target
    _fVel := DL_VM_ZERO;                        // 速度归零，从静止重新起算 / the velocity restarts from standstill
    _eState := E_DL_VMasterState.eIdle;         // 复位后回待机，由待机态按使能重判 / return to idle and let the enable decide the next phase
    IF NOT bError THEN
        eErr := 16#0004_01D8;                   // 信息级：相位复位已执行 / info: the phase reset was executed
    END_IF
END_IF

// 段 6｜斜坡与积分（故障拍与故障相均冻结：bError 或已处 eFault 皆不积分，修复前绝不带病复跑）
// segment 6, ramp and integration, frozen on a fault scan and inside the fault phase alike
IF (NOT bError) AND (_eState <> E_DL_VMasterState.eFault) THEN
    _fDtSec := DINT_TO_REAL(TIME_TO_DINT(tSample)) / DL_VM_MS_PER_S;    // 采样周期折算秒值 [s] / sample period in seconds
    _fMaxUp := fAccLimit * _fDtSec;             // 本拍允许上升量 [mm/s] / permitted increase of this scan
    _fMaxDn := fDecLimit * _fDtSec;             // 本拍允许下降量 [mm/s] / permitted decrease of this scan
    _fDiff := _fTarget - _fVel;                 // 目标与当前之差 [mm/s] / target minus current
    _fDelta := LIMIT(DL_VM_ZERO - _fMaxDn, _fDiff, _fMaxUp);    // 限幅后的增量 [mm/s]/ clipped increment [mm/s]
    IF ABS(_fDiff - _fDelta) > DL_VM_EPS THEN
        bLimited := TRUE;                       // 增量被截断，说明仍在斜坡 / the increment was clipped, the ramp is still active
    END_IF
    _fVel := _fVel + _fDelta;                   // 速度积分一格 / advance the velocity by one step
    IF _fDtSec > DL_VM_ZERO THEN
        fMasterAcc := _fDelta / _fDtSec;        // 本拍实际加速度，除子已判正 [mm/s²] / applied acceleration with a guarded divisor [mm/s²]
    END_IF
    _fPosL := _fPosL + REAL_TO_LREAL(_fVel * _fDtSec);    // 相位积分一格（步长先在 REAL 内算完再拓宽）[mm] / advance the phase by one step, the increment is computed in REAL and then widened [mm]

    // 精度门：越限即冻结并等调用方复位，绝不静默累计（凸轮错位的根源）
    // precision gate, freeze beyond the limit and wait for a reset instead of accumulating silently
    IF ABS(_fPosL) > DL_VM_POS_MAX THEN
        eErr := 16#0004_02EE;                   // 故障级：相位累计超 LREAL 有效精度 / fault: the phase accumulated beyond the effective LREAL precision
        bError := TRUE;                         // 置故障标志 / raise the fault flag
        _eState := E_DL_VMasterState.eFault;    // 转故障，相位冻结在当前值 / go to fault and freeze the phase at its current value
    END_IF
END_IF

// 段 7｜限幅信息码边沿发布：只在进入限幅的那一拍报，避免每拍刷屏
// segment 7, edge-published limiting info code, reported only on entry to limiting
IF bLimited AND (NOT _bLimitPrev) AND (NOT bError) THEN
    eErr := 16#0004_01D7;                       // 信息级：加速度限幅生效 / info: the acceleration limit is active
END_IF
_bLimitPrev := bLimited;                        // 更新限幅快照 / update the limiting snapshot

// 段 8｜状态机：只做可观测与转相判定，不承担斜坡职责（斜坡在段 6 已无条件算完）
// segment 8, the state machine only classifies and switches phases, the ramp itself lives in segment 6
IF NOT bError THEN
    CASE _eState OF
    E_DL_VMasterState.eIdle:
        // 待机：残速仍在段 6 递减；使能后按保持状态分相 / idle, the residual velocity still decays in segment 6
        IF bEnable AND bHold THEN
            _eState := E_DL_VMasterState.eHolding;  // 使能但要求保持 / enabled but holding
        ELSIF bEnable THEN
            _eState := E_DL_VMasterState.eRamping;  // 使能，进斜坡 / enabled, enter the ramp
        END_IF

    E_DL_VMasterState.eRamping:
        IF NOT bEnable THEN
            _eState := E_DL_VMasterState.eIdle;     // 失能，回待机按减速斜坡收尾 / disabled, finish through the deceleration ramp in idle
        ELSIF bHold THEN
            _eState := E_DL_VMasterState.eHolding;  // 转保持相 / enter the hold phase
        ELSIF ABS(_fTarget - _fVel) <= DL_VM_EPS THEN
            _eState := E_DL_VMasterState.eSteady;   // 达给定，进稳定相 / reached the setpoint
        END_IF

    E_DL_VMasterState.eSteady:
        IF NOT bEnable THEN
            _eState := E_DL_VMasterState.eIdle;     // 失能 / disabled
        ELSIF bHold THEN
            _eState := E_DL_VMasterState.eHolding;  // 转保持相 / enter the hold phase
        ELSIF ABS(_fTarget - _fVel) > DL_VM_EPS THEN
            _eState := E_DL_VMasterState.eRamping;  // 给定变了，重回斜坡 / the setpoint moved, ramp again
        END_IF

    E_DL_VMasterState.eHolding:
        IF NOT bEnable THEN
            _eState := E_DL_VMasterState.eIdle;     // 失能 / disabled
        ELSIF NOT bHold THEN
            _eState := E_DL_VMasterState.eRamping;  // 解除保持，重新向给定逼近 / hold released, ramp towards the setpoint again
        END_IF

    E_DL_VMasterState.eFault:
        // 故障退出：请求已撤且参数已修好；相位越精度门时还必须先复位（否则一拍后又越限）
        // fault exit, requires a withdrawn request and repaired parameters, plus a reset when the phase exceeded the precision gate
        IF (NOT bEnable) AND (NOT _bParamBad) THEN
            IF (ABS(_fPosL) <= DL_VM_POS_MAX) OR fbPhaseReset.Q THEN
                _eState := E_DL_VMasterState.eIdle;     // 允许回待机 / allowed back to idle
            END_IF
        END_IF

    ELSE
        // 非法状态兜底：绝不静默停在未知态 / illegal state fallback, never stay silently in an unknown state
        eErr := 16#0004_02EF;                   // 故障级：状态机落 ELSE / fault: the state machine fell into ELSE
        bError := TRUE;                         // 置故障标志 / raise the fault flag
        _eState := E_DL_VMasterState.eFault;    // 回故障态 / go to fault
    END_CASE
END_IF

// 段 9｜输出发布：相位只能从累加器读，绝不回读输出变量（R43 禁自反馈）
// segment 9, publish outputs; the phase is read from the accumulator only and never fed back from the output pin
fMasterPos := _fPosL;                           // 相位发布 [mm] / publish the phase [mm]
IF NOT bError THEN
    fMasterVel := _fVel;                        // 速度发布 [mm/s] / publish the velocity [mm/s]
END_IF
bReady := ((_eState = E_DL_VMasterState.eSteady)
           OR ((_eState = E_DL_VMasterState.eHolding) AND (ABS(_fVel) <= DL_VM_EPS))
           OR (_eState = E_DL_VMasterState.eIdle AND (ABS(_fVel) <= DL_VM_EPS)));    // 稳定或已停稳，主值可用 / settled or fully stopped, the master value may be consumed
bValid := NOT bError;                           // 输出可用 = 无故障级错误 / outputs are valid when no fault-level code is present
END_FUNCTION_BLOCK

(* ---- FC_DL_CamTableGenSeg.st ---- *)
(*
  ==================================================================
  组件名 Component  : FC_DL_CamTableGenSeg
  分类   Category   : DL_Motion
  复杂度 Complexity  : 中
  版本   Version    : 1.0.0
  功能   Purpose    : 凸轮表段型自动生成。按边界点（起点 / 终点）与点数生成
                      点列，段型三选一：线性 / 五次多项式（6u⁵-15u⁴+10u³）/
                      摆线（正弦修正单段位移式 u - sin(2πu)/(2π)）；生成后
                      做逐点单调性自检。供 CamTableValidate 前置使用。
  来源   Source     : t1-6-plcopen（凸轮族补口）
  溯源   Origin     : 段型位移表达式为公开凸轮设计教材内容（clean-room 整
                      理），生成与自检为自研实现，未复制 PLCopen 或任何厂商
                      私有库源码。
  平台   Platform   : 纯 IEC 61131-3，CODESYS / TwinCAT / InoProShop 通用
  分工声明 Split     : 与 DL_Motion 存量 FC_DL_CamTableValidate 分工——后者
                      验证既有凸轮表合法性，本件按段型生成点列供其前置；
                      本件不做电子凸轮耦合与主轴同步。
  作者   Author     : 道莅代码库 · PLC 编程专家（R58）
  ------------------------------------------------------------------
  功能说明  : 四段式防御（R45）：预置 → 非有限 / 点数域闸（钳位 2..64，信
              息级）→ 域内逐点生成（除子 nPoints-1 ≥ 1 已证）→ 单调性自检
              与结果非有限复检兜底。afTable 仅写 0..nPoints-1 槽位，其余槽
              位由调用方自行清理（本件不触碰，契约声明）。
  输出约定  : bOk = 生成受理；bClamped = 点数越域已钳位（信息级）；bMonoBad
              = 单调性自检失败（故障级，此时 bOk = FALSE）。
  修订记录  : 2026-11-21 v1.0.0 首次入库（R58 批 3 · 序号 12）
*)

(*-----------------------------------------------------------------------------
 * 枚举: E_DL_CamSegType（唯一属主 = 本文件，R67 全库唯一断言）
 * 含义: 凸轮表段型。
 *----------------------------------------------------------------------------*)
TYPE E_DL_CamSegType :
(
    eLinear  := 0, // 线性段 / the linear segment
    eQuintic := 1, // 五次多项式段 / the quintic segment
    eCycloid := 2  // 摆线段（正弦修正单段位移式）/ the cycloid segment, the sinusoid modified single segment form
);
END_TYPE

FUNCTION FC_DL_CamTableGenSeg : BOOL
VAR_INPUT
    eSegType  : E_DL_CamSegType; // 段型选择 [枚举] / the segment type selector
    fStartPos : LREAL; // 段起点位置 [工程单位] / the segment start position [engineering unit]
    fEndPos   : LREAL; // 段终点位置 [工程单位] / the segment end position [engineering unit]
    nPoints   : DINT;  // 生成点数 [个]，钳位 2..64 / the generated point count, clamped two through sixty four
END_VAR
VAR_IN_OUT
    afTable : ARRAY[0..63] OF LREAL; // 生成点列表 [工程单位]，仅写 0..nPoints-1 / the generated point list, only the first nPoints slots written
END_VAR
VAR_OUTPUT
    bOk      : BOOL; // 生成受理标志 [-] / the accepted flag
    bClamped : BOOL; // 点数越域钳位发生（信息级）[-] / a point count clamp happened, informational
    bMonoBad : BOOL; // 单调性自检失败（故障级）[-] / the monotony self check failed, fault grade
END_VAR
VAR
    lrSpan  : LREAL; // 段行程 [工程单位] / the segment span
    lrU     : LREAL; // 归一化进度 [无量纲] / the normalized progress
    lrS     : LREAL; // 段型形状因子 [无量纲] / the segment shape factor
    lrPos   : LREAL; // 点位置工作量 [工程单位] / the point position work value
    lrPrev  : LREAL; // 前点形状因子快照 [无量纲] / the previous shape factor snapshot
    lrSgn   : LREAL; // 方向号（+1 上行、-1 下行、0 平段）[无量纲] / the direction sign
    nPts    : DINT;  // 点数工作副本 [个] / the point count work copy
    nI      : DINT;  // 点遍历索引 [个] / the point loop index
    bBad    : BOOL;  // 故障级闸命中工作量 [-] / the fault gate work flag
END_VAR
VAR CONSTANT
    DL_CTS_NMAX   : DINT  := 64;                  // 点数上界 [个]，与数组容量一致 / the point bound, aligned with the array capacity
    DL_CTS_TWOPI  : LREAL := 6.283185307179586;   // 圆周率二倍（LREAL 精度字面量，R51）/ two pi at LREAL precision
END_VAR

// 段 1｜返回值与错误状态预置安全值（四段式第一段，R45）/ segment 1, preset the return and error states
FC_DL_CamTableGenSeg := FALSE; // 受理标志预置假 / preset the accepted flag false
bOk := FALSE; // 受理标志预置假 / preset the accepted flag false
bClamped := FALSE; // 钳位标志预置假 / preset the clamp flag false
bMonoBad := FALSE; // 单调标志预置假 / preset the mono flag false
bBad := FALSE; // 故障闸工作量预置假 / preset the fault work flag false

// 段 2｜非有限入参闸（起点终点双判据，R79）/ segment 2, the non finite input gate
IF (fStartPos <> fStartPos) OR ((fStartPos - fStartPos) <> (fStartPos - fStartPos)) THEN // 起点非有限 / a non finite start
    bBad := TRUE; // 置故障闸 / raise the fault gate
END_IF
IF (fEndPos <> fEndPos) OR ((fEndPos - fEndPos) <> (fEndPos - fEndPos)) THEN // 终点非有限 / a non finite end
    bBad := TRUE; // 置故障闸 / raise the fault gate
END_IF

// 段 3｜点数钳位（信息级，边界与数组容量一致，索引结构性安全）/ segment 3, the point count clamp
nPts := nPoints; // 装工作副本 / load the work copy
IF nPts < 2 THEN // 低于下界（单点无法构成段）/ below the floor
    nPts := 2; // 钳到 2 / clamp to two
    bClamped := TRUE; // 信息级钳位 / the informational clamp
ELSIF nPts > DL_CTS_NMAX THEN // 高于上界 / above the bound
    nPts := DL_CTS_NMAX; // 钳到容量 / clamp to the capacity
    bClamped := TRUE; // 信息级钳位 / the informational clamp
END_IF

// 段 4｜段型生成（除子 nPts-1 ≥ 1 已证；两极限自检见边界段）/ segment 4, the generation by the segment type
lrSpan := fEndPos - fStartPos; // 段行程 / the span
IF NOT bBad THEN // 无故障才生成 / generate only without a fault
    lrSgn := 0.0; // 方向号预置平段 / preset the sign zero
    IF lrSpan > 1.0E-12 THEN // 上行段 / an up segment
        lrSgn := 1.0; // 方向号置正 / the sign positive
    ELSIF lrSpan < -1.0E-12 THEN // 下行段 / a down segment
        lrSgn := -1.0; // 方向号置负 / the sign negative
    END_IF
    lrPrev := 0.0; // 前点因子快照预置零（首点因子恒 0）/ preset the previous snapshot
    FOR nI := 0 TO nPts - 1 DO // 逐点生成（固定界）/ the per point generation
        lrU := DINT_TO_LREAL(nI) / DINT_TO_LREAL(nPts - 1); // 归一化进度（除子已证 ≥1）/ the normalized progress
        CASE eSegType OF // 段型形状因子（边界点 s(0)=0 / s(1)=1 两极限自检成立）/ the shape factor, the both ends verified
        E_DL_CamSegType.eLinear: // 线性段 / the linear segment
            lrS := lrU; // 线性形状 / the linear shape
        E_DL_CamSegType.eQuintic: // 五次多项式段 / the quintic segment
            lrS := 10.0 * lrU * lrU * lrU - 15.0 * lrU * lrU * lrU * lrU + 6.0 * lrU * lrU * lrU * lrU * lrU; // 6u⁵-15u⁴+10u³ / the quintic form
        E_DL_CamSegType.eCycloid: // 摆线段（正弦修正单段位移式）/ the cycloid segment
            lrS := lrU - SIN(DL_CTS_TWOPI * lrU) / DL_CTS_TWOPI; // u - sin(2πu)/(2π) / the cycloidal form
        ELSE // 未知段型兜底（R128）/ the unknown segment fallback
            bBad := TRUE; // 置故障闸 / raise the fault gate
            lrS := 0.0; // 因子安全值 / the safe factor
        END_CASE
        lrPos := fStartPos + lrS * lrSpan; // 点位置 / the point position
        IF (lrPos <> lrPos) OR ((lrPos - lrPos) <> (lrPos - lrPos)) THEN // 点位置非有限（累乘溢出防御）/ a non finite point
            bBad := TRUE; // 置故障闸 / raise the fault gate
        END_IF
        IF NOT bBad THEN // 无故障才写表 / write the table only without a fault
            afTable[nI] := lrPos; // 写点（索引已证 < nPts ≤ 64）/ write the point
            IF nI > 0 THEN // 非首点做单调预检（逐点，最终判定在段 5）/ the per point mono pre check
                IF lrSgn > 0.0 THEN // 上行预检 / the up pre check
                    IF lrS < (lrPrev - 1.0E-12) THEN // 形状因子回落 / a shape dip
                        bMonoBad := TRUE; // 置单调失败 / raise the mono failure
                    END_IF
                ELSIF lrSgn < 0.0 THEN // 下行预检 / the down pre check
                    IF lrS > (lrPrev + 1.0E-12) THEN // 形状因子反弹 / a shape bounce
                        bMonoBad := TRUE; // 置单调失败 / raise the mono failure
                    END_IF
                END_IF // 平段（lrSgn = 0）无单调判据（两端点相等，逐点值恒等）
            END_IF
            lrPrev := lrS; // 快照推进 / advance the snapshot
        END_IF
    END_FOR
END_IF

// 段 5｜受理出口（单调失败为故障级，受理拒绝）/ segment 5, the acceptance outlet
IF bBad OR bMonoBad THEN // 故障或单调失败 / a fault or a mono failure
    FC_DL_CamTableGenSeg := FALSE; // 拒绝受理 / refuse the acceptance
ELSE // 正常受理 / the normal acceptance
    FC_DL_CamTableGenSeg := TRUE; // 受理 / accept
    bOk := TRUE; // 受理标志 / the accepted flag
END_IF
END_FUNCTION

(* ---- FC_DL_CamTableInterp.st ---- *)
(*==============================================================================
 * 组件名称 (Component)  : FC_DL_CamTableInterp
 * 溯源说明 (Provenance) : 道莅 clean-room 防御性实现（PLCopen 凸轮族深化）
 * 所属子库 (Sublibrary) : DL_Motion / CamProfile
 * 当前版本 (Version)    : 1.0.2
 * 兼容性   (Platform)   : CODESYS 3.5 / TwinCAT 3 / 汇川 InoProShop；
 *                         纯 IEC 61131-3（第 3 版），零标准库依赖
 * 组件分类 (Category)   : 函数（FUNCTION）· 凸轮表主轴位置线性插值（无状态纯函数）
 * 功能一句话 (Summary)  : 按主轴位置在凸轮表线性插值取从轴位置，支持周期取模。
 * 修复记录 (Fix)        : R75 解 VLA 透传（E037），增显式点数字段：
 *                         增入参 uPointCnt（1..200，内部钳位 [2,200]），
 *                         aCam 形参由 ARRAY[*] 改为固定上界 ARRAY[1..200]，
 *                         全部循环与下标以钳位后点数为界（调用方
 *                         FB_DL_CamOverrideTrim 已同步适配 v1.0.1）。
 * 边界与安全 (Boundary) : ①表点数钳位后 < 2 不可能，表非法仅由未升序/周期
 *                         非正触发；uPointCnt 越域静默钳位（本函数无信息码通道，
 *                         越域由调用方自行判码）；
 *                         ②主轴位置 NaN → 位置非法码；
 *                         ③非周期模式界外钳端点并 bInRange=FALSE；
 *                         ④周期模式先取模再插值，周期非正非法码；
 *                         ⑤纯函数：每个输出在全部路径（含提前返回）赋值。
 * 错误码    : 16#0004_0315 凸轮表非法（未升序或周期非正）——故障级
 *             16#0004_0316 主轴位置 NaN——故障级
 *             16#0004_0317 保留禁用（不得挪用，本件零赋值）
 * 码位总账  : 16#0004_0315 用 ｜ 16#0004_0316 用 ｜ 16#0004_0317 预留
 * 修改记录  : v1.0.0 R26 初版
 *             v1.0.1 R26 终审修复：周期参数补非有限闸——fPeriod=NaN 时
 *             `fPeriod <= 0.0` 判 FALSE 守卫穿透，NaN 经取模扩散至从轴输出
 *             v1.0.2 R75 显式点数字段修复：解 VLA 透传（E037），aCam 固定
 *             上界 ARRAY[1..200]，uPointCnt 钳位 [2,200]，下标改 1 基
 *==============================================================================*)
TYPE ST_DL_CamPoint :
STRUCT
    fMaster : LREAL; // 主轴位置锚点 [mm] / Master position anchor [mm]
    fSlave  : LREAL; // 从轴位置锚点 [mm] / Slave position anchor [mm]
END_STRUCT
END_TYPE

FUNCTION FC_DL_CamTableInterp : BOOL
VAR_INPUT
    fMasterPos : LREAL;               // 主轴当前位置 [mm] / Current master position [mm]
    bPeriodic  : BOOL;                // 周期模式使能 [-] / Periodic mode enable
    fPeriod    : LREAL;               // 周期模式主轴周期 [mm] / Master period [mm]
    uPointCnt  : UINT;                // 凸轮表有效点数，内部钳位 [2,200] [点] / Valid table point count, clamped internally
END_VAR
VAR_IN_OUT
    aCam : ARRAY[1..200] OF ST_DL_CamPoint; // 凸轮表（固定上界，须按 fMaster 升序且下标 1..uPointCnt 有效）/ Cam table, fixed bound, ascending over 1..uPointCnt
END_VAR
VAR_OUTPUT
    fSlavePos : LREAL;                // 从轴位置输出 [mm] / Slave position output [mm]
    bInRange  : BOOL;                 // 主轴位置在表界内 [-] / Master within table range
    eErr      : UDINT;                // 本周期错误码，0=无错 / Error code this cycle, 0 = none
END_VAR
VAR
    nPts    : INT;                    // 钳位后表点数 [点] / Clamped table point count
    i       : INT;                    // 分段搜索游标 / Segment search cursor
    fPos    : LREAL;                  // 插值用主轴位置（取模后）[mm] / Master position used for interpolation
    fDen    : LREAL;                  // 段宽（前判零）[mm] / Segment width, zero-guarded
    fRatio  : LREAL;                  // 段内插值比例 [-] / Interpolation ratio
    bTableOk: BOOL;                   // 表合法性 [-] / Table legality
END_VAR

// ---------- 全路径赋值缺省 ----------
fSlavePos := 0.0;
bInRange  := FALSE;
eErr      := 0;
FC_DL_CamTableInterp := TRUE; // 返回值：TRUE=已执行 / Result: TRUE = executed

// ---------- 点数钳位 [2, 200]（R75 显式点数字段口径） ----------
nPts := UINT_TO_INT(uPointCnt);               // 点数转整型 / Point count to INT
IF nPts < 2 THEN
    nPts := 2;                                // 下限钳 2（至少两点） / Clamp lower to 2
END_IF
IF nPts > 200 THEN
    nPts := 200;                              // 上限钳 200（数组容量） / Clamp upper to 200
END_IF

// ---------- 表防御：单调性（点数钳位后恒 >= 2） ----------
bTableOk := TRUE;                             // 合法性初值 / Legality init
FOR i := 1 TO nPts - 1 DO
    IF NOT (aCam[i].fMaster < aCam[i + 1].fMaster) THEN
        bTableOk := FALSE;                    // 严格升序被破坏 / Order violated
    END_IF
END_FOR
IF bPeriodic AND ((fPeriod <= 0.0) OR (fPeriod <> fPeriod)) THEN
    bTableOk := FALSE;                        // 周期非正或非有限视同表非法 / Non-positive or non-finite period illegal
END_IF
IF NOT bTableOk THEN
    eErr := 16#0004_0315;                     // 表非法码 / Illegal table code
    RETURN;                                   // 提前返回：输出已全赋值 / Early return, outputs assigned
END_IF

// ---------- 主轴位置 NaN 拦截 ----------
IF fMasterPos <> fMasterPos THEN
    eErr := 16#0004_0316;                     // 位置非法码 / Illegal position code
    RETURN;                                   // 提前返回：输出已全赋值 / Early return, outputs assigned
END_IF

// ---------- 周期模式取模（分母前判零） ----------
fPos := fMasterPos;
IF bPeriodic THEN
    fPos := fMasterPos - DINT_TO_LREAL(TRUNC(fMasterPos / fPeriod)) * fPeriod; // 取模 / Modulo
    IF fPos < 0.0 THEN
        fPos := fPos + fPeriod;               // 负余数钳回正域 / Negative remainder fixed
    END_IF
END_IF

// ---------- 界外处理：非周期钳端点并置界外标志 ----------
IF fPos <= aCam[1].fMaster THEN               // 界下判定（1 基下标）/ Below-range check
    fSlavePos := aCam[1].fSlave;              // 界下钳首点 / Clamp to first point
    IF fPos < aCam[1].fMaster THEN
        bInRange := FALSE;                    // 严格界外标志 / Strictly out of range
    ELSE
        bInRange := TRUE;                     // 恰在首点界内 / Exactly at first point
    END_IF
    RETURN;
END_IF
IF fPos >= aCam[nPts].fMaster THEN            // 界上判定 / Above-range check
    fSlavePos := aCam[nPts].fSlave;           // 界上钳末点 / Clamp to last point
    IF fPos > aCam[nPts].fMaster THEN
        bInRange := FALSE;
    ELSE
        bInRange := TRUE;
    END_IF
    RETURN;
END_IF

// ---------- 段定位与线性插值（i ∈ [1, nPts-1]，下标 i/i+1 均有界） ----------
bInRange := TRUE;                             // 界内插值 / In-range interpolation
i := 1;
WHILE (i < nPts - 1) AND (fPos > aCam[i + 1].fMaster) DO
    i := i + 1;                               // 定位所在段 / Locate segment
END_WHILE
fDen := aCam[i + 1].fMaster - aCam[i].fMaster; // 段宽 / Segment width
IF fDen > 0.0 THEN
    fRatio := (fPos - aCam[i].fMaster) / fDen; // 除法前判零 / Zero-guarded divide
    fSlavePos := aCam[i].fSlave + fRatio * (aCam[i + 1].fSlave - aCam[i].fSlave); // 插值 / Interpolate
ELSE
    fSlavePos := aCam[i].fSlave;              // 零段宽防御取左点 / Zero-width defensive
END_IF

END_FUNCTION

(* ---- FC_DL_WebGuideOffsetCalc.st ---- *)
(*
  Component : FC_DL_WebGuideOffsetCalc
  Category  : DL_Motion
  Function  : 纠偏偏移量计算：边缘模式取单侧偏差，中心模式取双传感器均值差，输出带符号偏移
  Complexity: C2
  开源溯源 : DLF 内部原创（R94 族模板派生）；参考语义来源见 SOURCE_HUNTING_MATRIX.md
  规则遵从 : R1-R16
  契约     : 输入 eMode 检测模式枚举、rEdgeLeftMm 左侧传感器距离 [mm]、rEdgeRightMm 右侧传感器距离 [mm]、
             rSensorSpanMm 两传感器安装跨距 [mm]、rCenterRefMm 目标中心（跨距中点为零点） [mm]；
             输出 rOffsetMm 带符号偏移（正=卷材偏右） [mm]、rCenterPosMm 卷材中心位置 [mm]、
             xValid 有效标志、nFaultCode 故障码。
  边界     : 边缘模式只用左侧传感器，中心位置 = 左侧距离；中心模式中心位置 = (左距离 + (跨距 − 右距离))/2，
             跨距须 >1.0E-6 [mm]；偏移为带符号量，不做钳位（符号即纠偏方向，钳位会反转方向）。
  码位     : 9801 输入非有限（故障级）；9802 跨距越域（故障级）；9803 模式枚举未知（故障级）。
*)
TYPE E_DL_WebGuideMode :
(
    eEdge   := 0,    // 边缘模式：单侧传感器对边 EN: the edge mode using one side sensor
    eCenter := 1     // 中心模式：双传感器对中 EN: the center mode using two sensors
);
END_TYPE

FUNCTION FC_DL_WebGuideOffsetCalc : BOOL
VAR_INPUT
    eMode        : E_DL_WebGuideMode;   // 检测模式 [-] EN: the detection mode
    rEdgeLeftMm  : LREAL := 50.0;       // 左侧传感器到卷材边距离 [mm] EN: the distance from the left sensor to the web edge
    rEdgeRightMm : LREAL := 50.0;       // 右侧传感器到卷材边距离 [mm] EN: the distance from the right sensor to the web edge
    rSensorSpanMm: LREAL := 400.0;      // 两传感器安装跨距 [mm] EN: the mounting span between the two sensors
    rCenterRefMm : LREAL := 200.0;      // 目标中心位置（相对左传感器） [mm] EN: the target center position relative to the left sensor
END_VAR
VAR_OUTPUT
    rOffsetMm    : LREAL;               // 带符号偏移，正表示卷材偏右 [mm] EN: the signed offset, positive means the web is to the right
    rCenterPosMm : LREAL;               // 卷材中心实测位置 [mm] EN: the measured web center position
    xValid       : BOOL;                // 输出可信标志 EN: the outputs are valid
    nFaultCode   : INT;                 // 0=无故障 9801=输入非有限 9802=跨距越域 9803=模式未知 EN: zero none, 9801 non finite, 9802 span out of range, 9803 unknown mode
END_VAR
VAR
    xFinAll  : BOOL;                    // 四个浮点入参有限 EN: the four floating inputs are finite
    rCenter  : LREAL;                   // 中心位置中间值 [mm] EN: the interim center position
    rOff     : LREAL;                   // 偏移中间值 [mm] EN: the interim offset
END_VAR
VAR CONSTANT
    DL_WGO_Z     : LREAL := 0.0;        // 浮点零常量 EN: the floating point zero constant
    DL_WGO_TWO   : LREAL := 2.0;        // 双侧平均系数 EN: the two sided averaging factor
    DL_WGO_MIN   : LREAL := 1.0E-6;     // 跨距下限 [mm] EN: the lower bound of the span
    DL_WGO_C_BAD : INT := 9801;         // 输入非有限 EN: a non finite input
    DL_WGO_C_SPAN: INT := 9802;         // 跨距越域 EN: the span is out of range
    DL_WGO_C_MODE: INT := 9803;         // 模式枚举未知 EN: the mode is unknown
END_VAR

// 段1｜出口预置
FC_DL_WebGuideOffsetCalc := FALSE;   // 返回值预置假 EN: preset the return value to false
rOffsetMm := DL_WGO_Z;               // 偏移预置零 [mm] EN: preset the offset to zero
rCenterPosMm := DL_WGO_Z;            // 中心位置预置零 [mm] EN: preset the center position to zero
xValid := FALSE;                     // 有效标志预置假 EN: preset the validity flag to false
nFaultCode := 0;                     // 故障码预置零 EN: preset the fault code to zero

// 段2｜非有限闸：四浮点入参全列（跨距与目标中心参与换算，漏则偏移静默失效）
xFinAll := (rEdgeLeftMm = rEdgeLeftMm) AND ((rEdgeLeftMm - rEdgeLeftMm) = DL_WGO_Z)
        AND (rEdgeRightMm = rEdgeRightMm) AND ((rEdgeRightMm - rEdgeRightMm) = DL_WGO_Z)
        AND (rSensorSpanMm = rSensorSpanMm) AND ((rSensorSpanMm - rSensorSpanMm) = DL_WGO_Z)
        AND (rCenterRefMm = rCenterRefMm) AND ((rCenterRefMm - rCenterRefMm) = DL_WGO_Z);   // 四输入有限性 EN: the finiteness of all four inputs
IF NOT xFinAll THEN                                                                          // 非有限出口 EN: leave early on a non finite input
    nFaultCode := DL_WGO_C_BAD;                                                              // 非有限码 EN: the non finite code
    RETURN;                                                                                  // 早退 EN: return early
END_IF

// 段3｜域闸：跨距必须足够大，否则中心模式分母退化
IF ABS(rSensorSpanMm) < DL_WGO_MIN THEN                                                      // 跨距下限 EN: the span magnitude gate
    nFaultCode := DL_WGO_C_SPAN;                                                             // 跨距越域码 EN: the span code
    RETURN;                                                                                  // 早退 EN: return early
END_IF

// 段4｜模式分派：ENUM + CASE 且 ELSE 兜底
CASE eMode OF
    E_DL_WebGuideMode.eEdge:
        rCenter := rEdgeLeftMm;                                                              // 边缘模式：左边缘即位置 [mm] EN: the edge mode uses the left edge as the position
    E_DL_WebGuideMode.eCenter:
        rCenter := (rEdgeLeftMm + (rSensorSpanMm - rEdgeRightMm)) / DL_WGO_TWO;              // 中心模式：两边中点 [mm] EN: the center mode averages both edges
ELSE
    nFaultCode := DL_WGO_C_MODE;                                                             // 未知模式码 EN: the unknown mode code
    RETURN;                                                                                  // 早退 EN: return early
END_CASE

// 段5｜偏移 = 实测中心 − 目标中心（符号保留方向）
rOff := rCenter - rCenterRefMm;                                                              // 带符号偏移 [mm] EN: the signed offset
IF (rOff <> rOff) OR (rCenter <> rCenter) THEN                                               // 结果复检 EN: recheck the result
    nFaultCode := DL_WGO_C_BAD;                                                              // 复检失败码 EN: the recheck failure code
    RETURN;                                                                                  // 早退，出口保持零哨兵 EN: return early with the zero sentinels
END_IF
rOffsetMm := rOff;                                                                           // 偏移出口 [mm] EN: the offset output
rCenterPosMm := rCenter;                                                                     // 中心位置出口 [mm] EN: the center position output
xValid := TRUE;                                                                              // 结果可信 EN: the results are valid
FC_DL_WebGuideOffsetCalc := TRUE;                                                            // 返回真 EN: return true
END_FUNCTION

(* ---- I_DL_ExternalEncoder.st ---- *)
(*==============================================================================
 * 组件名称 (Component)  : I_DL_ExternalEncoder
 * 所属子库 (Sublibrary) : DL_Motion
 * 前缀     (Prefix)     : I_DL_
 * 当前版本 (Version)    : 1.0.0
 * 兼容性   (Platform)   : CODESYS 3.5 / TwinCAT 3 / 汇川 InoProShop / Schneider
 *                         Machine Expert；纯 IEC 61131-3（第 3 版）接口语法，
 *                         无任何厂商方言、无标准库依赖（纯契约件）
 * 作者     (Author)     : 道莅代码库 · PLC编程专家（R31）
 * 开源溯源 (Origin)     : 外部编码器只读位置源公开契约语义（T1-6 外部编码器
 *                         族开族件），道莅 clean-room 防御性实现，
 *                         未复制任何外部源码行
 * 功能描述 (Function)   : 外部编码器契约接口，定义「外部编码器 = 只读位置源」
 *                         最小契约：三条只读属性回答"在哪、多快、可信吗"，
 *                         一个采样方法输出单拍一致快照（位置 + 速度 + 时戳
 *                         同拍锁定），一个复位方法。核心语义写死：外部编码器
 *                         不可被驱动，本接口无任何命令方向属性或方法。
 * 接口结构 (Contract)   : 1 属性：fPos / fVel / bValid 共 3 条，全部只读 GET；
 *                         2 方法：Sample / Reset 共 2 个（满足方法不超过 6 个
 *                         的拆分红线）；3 结构体：ST_DL_EncSnapshot 随本文件
 *                         发布，全库唯一属主为本文件。
 * 实现纪律 (Discipline) : 实现块不得在本接口后挂写方法或属性——外部编码器
 *                         不可被驱动是该族的编译期表达，任何写入型成员都
 *                         会破坏「只读位置源」契约。bValid=FALSE 的具体解释
 *                         （断线/超时/未标定）由实现块自行定义。
 * 码位     (Codes)      : 纯契约件无执行体，无错误码出口；段 16#0004_0063~0066
 *                         为本契约预留 4 槽（规格 §3 分配），实现块的错误码
 *                         不得挪用该段（段位隔离，防跨件码冲突）。
 * 边界防错 (Boundary)   : 1 接口不声明变量段（IEC 接口只允许属性与方法）；
 *                         2 Sample 的快照输出以 IN-OUT 引用传递承载规格的
 *                         OUT 语义（可移植性裁定，全平台语法一致）；
 *                         3 单拍一致快照由实现块保证：一次 Sample 调用内
 *                         位置、速度、时戳必须同拍锁定，不得跨拍拼装。
 * 修订历史 (Revision)   : 2026-11-18 v1.0.0 首版入库（R31 · 阶段三 · 序 5）
 *==============================================================================*)

(*------------------------------------------------------------------------------
 * 结构体: ST_DL_EncSnapshot（归属本接口，同文件发布，全库唯一属主）
 * 含义: 外部编码器单拍一致快照。实现块在一次 Sample 调用内同拍锁定全部字段。
 *----------------------------------------------------------------------------*)
TYPE ST_DL_EncSnapshot :
STRUCT
    fPos    : LREAL := 0.0;   // 快照位置 [毫米] / Snapshot position [mm]
    fVel    : LREAL := 0.0;   // 快照速度 [毫米每秒] / Snapshot velocity [mm per s]
    tStamp  : TIME  := T#0MS; // 快照时戳：实现块自填的采样时标 [毫秒] / Snapshot timestamp [ms]
    bValid  : BOOL  := FALSE; // 快照有效标志：实现块解释失效原因 / Snapshot validity, reason per implementation
END_STRUCT
END_TYPE

(*------------------------------------------------------------------------------
 * 接口: I_DL_ExternalEncoder
 * 契约结构: 属性（只读 GET，3 条）+ 方法（2 个）两段式。
 *----------------------------------------------------------------------------*)
INTERFACE I_DL_ExternalEncoder

// ---- 属性段（全部只读 GET，共 3 条）----------------------------------------

PROPERTY fPos   : LREAL   // 当前位置 [毫米] / Current position [mm]
END_PROPERTY
PROPERTY fVel   : LREAL   // 当前速度 [毫米每秒] / Current velocity [mm per s]
END_PROPERTY
PROPERTY bValid : BOOL    // 当前数据可信标志 / Current data validity flag
END_PROPERTY

// ---- 方法段（共 2 个）-------------------------------------------------------

// Sample：取单拍一致快照，成功返回 TRUE 且 stSnap 各字段同拍锁定；
// 失败返回 FALSE，stSnap 内容由实现块决定（约定不清写，调用方自行保持旧值）。
METHOD Sample : BOOL
VAR_IN_OUT
    stSnap : ST_DL_EncSnapshot; // 快照出参（IN-OUT 引用承载 OUT 语义）/ Snapshot output via in-out reference
END_VAR

// Reset：复位实现块内部采样历史（首扫同步标志、失效计数等），始终返回 TRUE。
// 只清采样历史，不清物理编码器状态（清零/回零属驱动层职责，不在本契约内）。
    END_METHOD

METHOD Reset : BOOL

    END_METHOD
END_INTERFACE

(* ---- FC_DL_AckermannSteerPairCalc.st ---- *)
// FC_DL_AckermannSteerPairCalc v1.0.0
// 开源溯源：clean-room 自研（族 DL_Motion，ST 生态实测 0 命中，无外部代码引入）
(*
  功能: 阿克曼内外轮角：R = L/tan|δ|，δin = ATAN(L/(R − T/2))，δout = ATAN(L/(R + T/2))，
        按 δ 符号回填正负；|δ| < 1e-4 视为直行，两轮同角（避开 tan 近零除爆）。
  邻件/码位: 与 FC_DL_StanleySteerAngleCalc 串联，把中心轮转角展开为内外轮；
             16#0002_9206 = 非有限、轴距轮距非正或转向几何不可达拒收。
*)
FUNCTION FC_DL_AckermannSteerPairCalc : REAL
VAR_INPUT
    fSteerCenter : REAL := 0.0;     // 中心轮转角 δ [rad]，右转为正 / Center steer angle [rad]
    fWheelBase   : REAL := 2.5;     // 轴距 L [m]，域 > 0 / Wheel base [m]
    fTrackWidth  : REAL := 1.5;     // 轮距 T [m]，域 > 0 / Track width [m]
END_VAR
VAR_OUTPUT
    fSteerInner : REAL;             // 内轮转角 [rad]，与中心同号 / Inner angle [rad]
    fSteerOuter : REAL;             // 外轮转角 [rad]，与中心同号 / Outer angle [rad]
    bValid      : BOOL;             // 结果有效回执 [-] / Result validity receipt
    uErrorId    : UDINT;            // 事件码，0 = 无事件 / Event code
END_VAR
VAR
    fAbsDelta : REAL := 0.0;        // 中心转角绝对值 [rad] / Absolute center angle [rad]
    fRadius   : REAL := 0.0;        // 后轴中心转弯半径 R [m] / Turning radius [m]
    fHalfTrk  : REAL := 0.0;        // 半轮距 T/2 [m] / Half track width [m]
    fInner    : REAL := 0.0;        // 内轮转角幅值 [rad] / Inner angle magnitude [rad]
    fOuter    : REAL := 0.0;        // 外轮转角幅值 [rad] / Outer angle magnitude [rad]
END_VAR
// 段 0：全路径出口安全缺省（内外轮零 = 直行）/ Safe defaults, zero angles mean straight
fSteerInner := 0.0;             // 内轮转角缺省零 / Inner angle default zero
fSteerOuter := 0.0;             // 外轮转角缺省零 / Outer angle default zero
bValid := FALSE;                // 有效回执预清 / Validity preset clear
uErrorId := 16#0000;            // 事件码预清 / Event code preset clear
FC_DL_AckermannSteerPairCalc := 0.0;    // 返回值缺省零（镜像内轮）/ Return default zero
// 段 1：非有限闸（三入参全枚举）/ Non-finite gate over all inputs
IF (fSteerCenter <> fSteerCenter) OR (fWheelBase <> fWheelBase) OR (fTrackWidth <> fTrackWidth)
   OR (ABS(fSteerCenter) >= 3.0E38) OR (ABS(fWheelBase) >= 3.0E38) OR (ABS(fTrackWidth) >= 3.0E38) THEN
    uErrorId := 16#0002_9206;   // 入参非有限拒收 / Non-finite input reject
    RETURN;
END_IF
// 段 2：域闸（轴距轮距为正 + 直行快通道 + 转向几何可达）/ Domain gate
IF (fWheelBase <= 1.0E-6) OR (fTrackWidth <= 1.0E-6) THEN
    uErrorId := 16#0002_9206;   // 轴距或轮距非正 / Non-positive base or track
    RETURN;
END_IF
fAbsDelta := fSteerCenter;                                      // 先直取中心转角 / Take center angle
IF fAbsDelta < 0.0 THEN
    fAbsDelta := -fAbsDelta;                                    // 取绝对值 / Absolute value
END_IF
IF fAbsDelta < 1.0E-4 THEN                                       // 直行快通道 / Straight fast path
    bValid := TRUE;                                             // 直行亦为有效解 / Straight is valid
    RETURN;                                                     // 两轮同角零已由段 0 给出 / Both zero from stage 0
END_IF
fHalfTrk := fTrackWidth / 2.0;                                  // 半轮距 / Half track
fRadius := fWheelBase / TAN(fAbsDelta);                         // R = L/tan|δ| [m] / Turning radius
IF (fRadius - fHalfTrk) <= 1.0E-6 THEN
    uErrorId := 16#0002_9206;   // 内轮半径非正，几何不可达 / Geometry unreachable
    RETURN;
END_IF
// 段 3：主计算（内外轮幅值 + 符号回填）/ Main computation
fInner := ATAN(fWheelBase / (fRadius - fHalfTrk));               // 内轮幅值 / Inner magnitude
fOuter := ATAN(fWheelBase / (fRadius + fHalfTrk));               // 外轮幅值 / Outer magnitude
fSteerInner := fInner;                                          // 先按右转（正）落值 / Assume right turn first
fSteerOuter := fOuter;                                          // 先按右转（正）落值 / Assume right turn first
IF fSteerCenter < 0.0 THEN
    fSteerInner := -fInner;                                     // 左转回填负号 / Negative for left turn
    fSteerOuter := -fOuter;                                     // 左转回填负号 / Negative for left turn
END_IF
// 段 4：出口闸（双角非有限复核 + 内大于外几何自检）/ Outlet gate
IF (fSteerInner <> fSteerInner) OR (fSteerOuter <> fSteerOuter)
   OR (ABS(fSteerInner) >= 3.0E38) OR (ABS(fSteerOuter) >= 3.0E38)
   OR (ABS(fSteerInner) < ABS(fSteerOuter)) THEN
    fSteerInner := 0.0;         // 复核失败回缺省 / Fallback on recheck failure
    fSteerOuter := 0.0;         // 复核失败回缺省 / Fallback on recheck failure
    uErrorId := 16#0002_9206;   // 出口复核拒收 / Output recheck reject
    RETURN;
END_IF
bValid := TRUE;                 // 有效回执 / Validity receipt
FC_DL_AckermannSteerPairCalc := fSteerInner;    // 返回值镜像内轮 / Return mirrors inner angle
END_FUNCTION

(* ---- FC_DL_AgvChargeDockAlignCalc.st ---- *)
// FC_DL_AgvChargeDockAlignCalc v1.0.0
// 开源溯源：clean-room 自研（族 DL_Motion，ST 生态实测 0 命中，无外部代码引入）
(*
  功能: 充电桩对桩对齐律：bAligned = (|Δy| ≤ tolY) AND (|Δa| ≤ tolA)；
        v = MIN(0.15, 0.3·dist)（dist 负则 0）；ω = 1.5·Δa 限幅 ±0.4 rad/s；
        已对齐强制零速零转（防贴桩抖动）。
  邻件/码位: 与 FC_DL_AgvSpeedLimitProfileCalc 分工（末端对桩 vs 巡航限速）；
             DOCK 相超时由 FB_DL_AgvPathTrackSeq 处理；16#0002_9209 = 域外或非有限拒收。
*)
FUNCTION FC_DL_AgvChargeDockAlignCalc : REAL
VAR_INPUT
    fOffsetY   : REAL := 0.0;       // 横向偏差 Δy [m]，左正 / Lateral offset [m]
    fAngleErr  : REAL := 0.0;       // 角度偏差 Δa [rad]，左正 / Angular error [rad]
    fDist      : REAL := 1.0;       // 到桩距离 [m] / Distance to dock [m]
    fAlignTolY : REAL := 0.02;      // 横向容差 [m]，负值归零 / Lateral tolerance [m]
    fAlignTolA : REAL := 0.03;      // 角度容差 [rad]，负值归零 / Angular tolerance [rad]
END_VAR
VAR_OUTPUT
    fSpeedCmd   : REAL;             // 前进速度指令 [m/s] / Forward speed command [m/s]
    fYawRateCmd : REAL;             // 转向角速度指令 [rad/s] / Yaw rate command [rad/s]
    bAligned    : BOOL;             // 对齐到位标志 [-] / Alignment reached flag
    bValid      : BOOL;             // 结果有效回执 [-] / Result validity receipt
    uErrorId    : UDINT;            // 事件码，0 = 无事件 / Event code
END_VAR
VAR
    fTolY   : REAL := 0.0;          // 生效横向容差 [m] / Effective lateral tolerance [m]
    fTolA   : REAL := 0.0;          // 生效角度容差 [rad] / Effective angular tolerance [rad]
    fYawRaw : REAL := 0.0;          // 未限幅转向指令 [rad/s] / Unsaturated yaw [rad/s]
END_VAR
// 段 0：全路径出口安全缺省（零速零转）/ Safe defaults, zero speed and zero yaw
fSpeedCmd := 0.0;               // 速度指令缺省零 / Speed command default zero
fYawRateCmd := 0.0;             // 转向指令缺省零 / Yaw command default zero
bAligned := FALSE;              // 对齐标志预清 / Alignment preset clear
bValid := FALSE;                // 有效回执预清 / Validity preset clear
uErrorId := 16#0000;            // 事件码预清 / Event code preset clear
FC_DL_AgvChargeDockAlignCalc := 0.0;    // 返回值缺省零（镜像速度）/ Return default zero
// 段 1：非有限闸（五入参全枚举）/ Non-finite gate over all inputs
IF (fOffsetY <> fOffsetY) OR (fAngleErr <> fAngleErr) OR (fDist <> fDist)
   OR (fAlignTolY <> fAlignTolY) OR (fAlignTolA <> fAlignTolA)
   OR (ABS(fOffsetY) >= 3.0E38) OR (ABS(fAngleErr) >= 3.0E38) OR (ABS(fDist) >= 3.0E38)
   OR (ABS(fAlignTolY) >= 3.0E38) OR (ABS(fAlignTolA) >= 3.0E38) THEN
    uErrorId := 16#0002_9209;   // 入参非有限拒收 / Non-finite input reject
    RETURN;
END_IF
// 段 2：域闸（容差负值归零，防误判永远对齐）/ Domain gate on tolerances
fTolY := fAlignTolY;                                            // 横向容差直取 / Take tolerance
IF fTolY < 0.0 THEN
    fTolY := 0.0;                                               // 负容差归零 / Clamp negative
END_IF
fTolA := fAlignTolA;                                            // 角度容差直取 / Take tolerance
IF fTolA < 0.0 THEN
    fTolA := 0.0;                                               // 负容差归零 / Clamp negative
END_IF
// 段 3：主计算（对齐判定 + 速度/转向生成）/ Main computation
IF (ABS(fOffsetY) <= fTolY) AND (ABS(fAngleErr) <= fTolA) THEN
    bAligned := TRUE;                                           // 双容差内判对齐 / Aligned
END_IF
IF NOT bAligned THEN
    IF fDist > 0.0 THEN
        fSpeedCmd := 0.3 * fDist;                               // 距离比例降速 / Distance proportional speed
        IF fSpeedCmd > 0.15 THEN
            fSpeedCmd := 0.15;                                  // 限到对桩上限 / Clamp to docking ceiling
        END_IF
    END_IF
    fYawRaw := 1.5 * fAngleErr;                                 // 角度比例转向 / Angular proportional yaw
    IF fYawRaw > 0.4 THEN
        fYawRateCmd := 0.4;                                     // 上饱和 / Upper saturation
    ELSIF fYawRaw < -0.4 THEN
        fYawRateCmd := -0.4;                                    // 下饱和 / Lower saturation
    ELSE
        fYawRateCmd := fYawRaw;                                 // 未饱和直通 / Pass through
    END_IF
END_IF
// 段 4：出口闸（双指令非有限复核）/ Outlet gate
IF (fSpeedCmd <> fSpeedCmd) OR (fYawRateCmd <> fYawRateCmd)
   OR (ABS(fSpeedCmd) >= 3.0E38) OR (ABS(fYawRateCmd) >= 3.0E38) THEN
    fSpeedCmd := 0.0;           // 复核失败回零速 / Fallback to zero speed
    fYawRateCmd := 0.0;         // 复核失败回零转 / Fallback to zero yaw
    bAligned := FALSE;          // 复核失败撤对齐 / Clear alignment
    uErrorId := 16#0002_9209;   // 出口非有限拒收 / Output non-finite reject
    RETURN;
END_IF
bValid := TRUE;                 // 有效回执 / Validity receipt
FC_DL_AgvChargeDockAlignCalc := fSpeedCmd;      // 返回值镜像速度指令 / Return mirrors speed
END_FUNCTION

(* ---- FC_DL_AgvSpeedLimitProfileCalc.st ---- *)
// FC_DL_AgvSpeedLimitProfileCalc v1.0.0
// 开源溯源：clean-room 自研（族 DL_Motion，ST 生态实测 0 命中，无外部代码引入）
(*
  功能: 曲率自适应限速：|κ| < 1e-4 判直道并取车最大速度；弯道按侧向加速度约束
        v = SQRT(a_lat/|κ|)，再向车最大速度取小。
  邻件/码位: 与 FC_DL_PurePursuitCurvatureCalc 衔接（曲率→限速）；对桩末端由
             FC_DL_AgvChargeDockAlignCalc 处理；16#0002_9208 = 非有限或域外拒收。
*)
FUNCTION FC_DL_AgvSpeedLimitProfileCalc : REAL
VAR_INPUT
    fPathCurvature : REAL := 0.0;   // 路径曲率 κ [1/m] / Path curvature [1/m]
    fLatAccMax     : REAL := 0.5;   // 允许侧向加速度 [m/s²]，域 > 0 / Lateral acceleration [m/s^2]
    fSpeedMax      : REAL := 1.5;   // 车最大速度 [m/s]，域 > 0 / Vehicle max speed [m/s]
END_VAR
VAR_OUTPUT
    fSpeedLimit : REAL;             // 限速结果 [m/s] / Speed limit result [m/s]
    bStraight   : BOOL;             // 直道标志 [-] / Straight-path flag
    bValid      : BOOL;             // 结果有效回执 [-] / Result validity receipt
    uErrorId    : UDINT;            // 事件码，0 = 无事件 / Event code
END_VAR
VAR
    fAbsKappa : REAL := 0.0;        // 曲率绝对值 |κ| [1/m] / Absolute curvature [1/m]
END_VAR
// 段 0：全路径出口安全缺省（限速零 = 最保守）/ Safe defaults, zero limit is conservative
fSpeedLimit := 0.0;             // 限速缺省零 / Speed limit default zero
bStraight := FALSE;             // 直道标志预清 / Straight flag preset clear
bValid := FALSE;                // 有效回执预清 / Validity preset clear
uErrorId := 16#0000;            // 事件码预清 / Event code preset clear
FC_DL_AgvSpeedLimitProfileCalc := 0.0;  // 返回值缺省零 / Return default zero
// 段 1：非有限闸（三入参全枚举）/ Non-finite gate over all inputs
IF (fPathCurvature <> fPathCurvature) OR (fLatAccMax <> fLatAccMax) OR (fSpeedMax <> fSpeedMax)
   OR (ABS(fPathCurvature) >= 3.0E38) OR (ABS(fLatAccMax) >= 3.0E38) OR (ABS(fSpeedMax) >= 3.0E38) THEN
    uErrorId := 16#0002_9208;   // 入参非有限拒收 / Non-finite input reject
    RETURN;
END_IF
// 段 2：域闸（侧向加速度与车最大速度为正）/ Domain gate
IF (fLatAccMax <= 1.0E-6) OR (fSpeedMax <= 1.0E-6) THEN
    uErrorId := 16#0002_9208;   // 上限非正，限速不可解 / Non-positive bound
    RETURN;
END_IF
fAbsKappa := ABS(fPathCurvature);                               // 曲率绝对值 / Absolute curvature
// 段 3：主计算（直道快通道 / 弯道侧向加速度约束）/ Main computation
IF fAbsKappa < 1.0E-4 THEN
    fSpeedLimit := fSpeedMax;                                   // 直道取车最大速度 / Straight: max speed
    bStraight := TRUE;                                          // 置直道标志 / Set straight flag
ELSE
    fSpeedLimit := SQRT(fLatAccMax / fAbsKappa);                // v = sqrt(a_lat/|κ|) / Curve-limited speed
    IF fSpeedLimit > fSpeedMax THEN
        fSpeedLimit := fSpeedMax;                               // 向车最大速度取小 / Clamp to max
    END_IF
END_IF
// 段 4：出口闸（非有限复核 + 非负复核）/ Outlet gate
IF (fSpeedLimit <> fSpeedLimit) OR (ABS(fSpeedLimit) >= 3.0E38) OR (fSpeedLimit < 0.0) THEN
    fSpeedLimit := 0.0;         // 复核失败回零速 / Fallback to zero speed
    bStraight := FALSE;         // 复核失败撤直道标志 / Clear straight flag
    uErrorId := 16#0002_9208;   // 出口复核拒收 / Output recheck reject
    RETURN;
END_IF
bValid := TRUE;                 // 有效回执 / Validity receipt
FC_DL_AgvSpeedLimitProfileCalc := fSpeedLimit;  // 返回值镜像限速 / Return mirrors limit
END_FUNCTION

(* ---- FC_DL_ArcCenterOffsetCalc.st ---- *)
(* ============================================================
   DL_Motion / FC_DL_ArcCenterOffsetCalc ｜ v1.0.0 ｜ 2026-11-25
   功能：由起点/终点/半径反解圆心相对起点偏移 [mm]；bCcw=TRUE 取劣弧（垂距正），
         FALSE 取优弧（垂距负）。弦向量左法向 × 垂距 h 即偏移。
   边界：半径<半弦长 或 起终点重合 → uErrId=1；半径≤0 或非有限 → uErrId=2，
         且实值出口同拍写 0（N1：判据与出口同源，禁 NaN 直穿）
   依赖：仅 IEC 61131-3（SQRT / MAX） ｜ 溯源：DLF-A-RTCP（内部原创线）
   ============================================================ *)
FUNCTION FC_DL_ArcCenterOffsetCalc : BOOL
VAR_INPUT
    fX1       : LREAL;   // 起点 X 坐标 [mm] / Start point X in mm
    fY1       : LREAL;   // 起点 Y 坐标 [mm] / Start point Y in mm
    fX2       : LREAL;   // 终点 X 坐标 [mm] / End point X in mm
    fY2       : LREAL;   // 终点 Y 坐标 [mm] / End point Y in mm
    fRadiusMm : LREAL;   // 圆弧半径，有效域 > 0 [mm] / Arc radius, domain above zero
    bCcw      : BOOL;    // TRUE=劣弧（圆心在弦左）[-] / TRUE selects the minor arc
END_VAR
VAR_OUTPUT
    fDx    : LREAL;   // 圆心相对起点 X 偏移 [mm] / Center offset in X
    fDy    : LREAL;   // 圆心相对起点 Y 偏移 [mm] / Center offset in Y
    uErrId : UDINT;   // 出口码 0 正常 / 1 几何不可解 / 2 入参非法 [-] / Outlet code
    bOk    : BOOL;    // 结果可信标志，与返回值同源 [-] / Result trustworthy flag
END_VAR
VAR
    _fCx   : LREAL;  // 弦向量 X 分量 [mm] / Chord vector X component
    _fCy   : LREAL;  // 弦向量 Y 分量 [mm] / Chord vector Y component
    _fLen  : LREAL;  // 弦长 [mm] / Chord length
    _fHalf : LREAL;  // 半弦长 [mm] / Half chord length
    _fH    : LREAL;  // 圆心到弦中点垂距 [mm] / Perpendicular from chord midpoint to center
END_VAR
VAR CONSTANT
    DL_ARC_EPS : LREAL := 1.0E-9;  // 几何判零容差 [mm] / Geometric zero tolerance
END_VAR

(* 段 0：出口预置安全侧 + 非有限双判闸（NaN 自反 + Inf 差值自减，R79） *)
FC_DL_ArcCenterOffsetCalc := FALSE;
fDx := 0.0;  fDy := 0.0;  uErrId := 2;  bOk := FALSE;
IF (fX1 <> fX1) OR (fY1 <> fY1) OR (fX2 <> fX2) OR (fY2 <> fY2) OR (fRadiusMm <> fRadiusMm) THEN
    RETURN;                                          // NaN：判据与出口同源于原始入参（N1）
END_IF
IF ((fX1 - fX1) <> (fX1 - fX1)) OR ((fY1 - fY1) <> (fY1 - fY1))
   OR ((fX2 - fX2) <> (fX2 - fX2)) OR ((fY2 - fY2) <> (fY2 - fY2))
   OR ((fRadiusMm - fRadiusMm) <> (fRadiusMm - fRadiusMm)) THEN
    RETURN;                                          // ±Inf：半径 +Inf 会直穿到出口 ±Inf 并报码 0
END_IF

(* 段 1：弦向量、半弦长与退化判定 *)
_fCx := fX2 - fX1;  _fCy := fY2 - fY1;
_fLen := SQRT(_fCx * _fCx + _fCy * _fCy);
IF _fLen <> _fLen THEN RETURN; END_IF               // 弦长运算产生 NaN 的兜底（入参 Inf 已由段 0 拦截）
IF _fLen <= DL_ARC_EPS THEN uErrId := 1; RETURN; END_IF  // 起终点重合 / Coincident points
_fHalf := _fLen / 2.0;

(* 段 2：半径域闸与可解性 *)
IF fRadiusMm <= 0.0 THEN RETURN; END_IF
IF fRadiusMm < (_fHalf - DL_ARC_EPS) THEN uErrId := 1; RETURN; END_IF

(* 段 3：垂距与位移分量（劣弧取正、优弧取负） *)
_fH := SQRT(MAX(0.0, fRadiusMm * fRadiusMm - _fHalf * _fHalf));
IF bCcw THEN
    fDx := (_fCx / 2.0) + _fH * (0.0 - _fCy) / _fLen;
    fDy := (_fCy / 2.0) + _fH * _fCx / _fLen;
ELSE
    fDx := (_fCx / 2.0) - _fH * (0.0 - _fCy) / _fLen;
    fDy := (_fCy / 2.0) - _fH * _fCx / _fLen;
END_IF

(* 段 4：结果复检 + 单一出口裁决（N4：实值与 bOk 同源改写） *)
IF (fDx <> fDx) OR (fDy <> fDy)
   OR ((fDx - fDx) <> (fDx - fDx)) OR ((fDy - fDy) <> (fDy - fDy)) THEN
    fDx := 0.0;  fDy := 0.0;  uErrId := 2;  bOk := FALSE;  RETURN;
END_IF
uErrId := 0;  bOk := TRUE;  FC_DL_ArcCenterOffsetCalc := TRUE;
END_FUNCTION

(* ---- FC_DL_BeltLengthCalc.st ---- *)
// FC_DL_BeltLengthCalc v1.0.0
// 开源溯源：self-cleanroom / 公开公式（开口带传动节线长度）
(*
  道莅工业代码库 | DL_Motion | FC_DL_BeltLengthCalc
  版本: 1.0.0 | 日期: 2026-11-23 | 轮次: R75
  功能: 开口平带/同步带节线长度：L = 2C + π(D1+D2)/2 + (D2−D1)²/(4C)，
        中心距分母域闸；D1/D2 为两轮节圆直径，大小顺序不限（公式对称）
  邻件关系: 与 FurnaceBeltTension / FanBeltSlipDiag（带张力/打滑诊断）同族 ——
            差异点：张力/打滑件为运行状态诊断，本件为选型长度计算（设计域），
            码位独立（本件 16#0002_2801）
*)
FUNCTION FC_DL_BeltLengthCalc : REAL
VAR_INPUT
    fDia1    : REAL := 50.0;    // 轮 1 节圆直径 D1 [mm]，域 >= 0 / Pitch diameter pulley 1 [mm]
    fDia2    : REAL := 50.0;    // 轮 2 节圆直径 D2 [mm]，域 >= 0 / Pitch diameter pulley 2 [mm]
    fCenter  : REAL := 200.0;   // 中心距 C [mm]，域 > 0 / Center distance [mm]
    fEps     : REAL := 1.0E-6;  // 判零容差 [mm] / Zero tolerance [mm]
END_VAR
VAR_OUTPUT
    fBeltLength : REAL;         // 节线长度 L [mm] / Pitch line length [mm]
    bValid      : BOOL;         // 结果有效回执 [-] / Result validity receipt
    uErrorId    : UDINT;        // 事件码，0 = 无事件；16#0002_2801 = 域外拒收 / Event code
END_VAR

// —— 段 0：全路径缺省 —— //
fBeltLength := 0.0;             // 长度缺省零 / Length default zero
bValid := FALSE;                // 有效回执预清 / Validity preset
uErrorId := 16#0000;            // 事件码预清 / Event code preset
FC_DL_BeltLengthCalc := 0.0;    // 返回值缺省零（镜像长度）/ Return default mirrors length

// —— 段 1：非有限闸 —— //
IF (fDia1 <> fDia1) OR (fDia2 <> fDia2) OR (fCenter <> fCenter)
   OR (ABS(fDia1) >= 3.0E38) OR (ABS(fDia2) >= 3.0E38) OR (ABS(fCenter) >= 3.0E38) THEN
    uErrorId := 16#0002_2801;   // 输入非有限拒收 / Non-finite reject
    RETURN;
END_IF

// —— 段 2：域闸（直径非负 + 中心距正数防零，R4） —— //
IF (fDia1 < 0.0) OR (fDia2 < 0.0) OR (fCenter < fEps) THEN
    uErrorId := 16#0002_2801;   // 信息级：直径为负或中心距近零（分母为零风险）/ Info level: domain violation
    RETURN;                     // 不计算返回 / Return without computation
END_IF

// —— 段 3：主计算（分母已过闸，公式对 D1/D2 对称） —— //
fBeltLength := 2.0 * fCenter
             + 3.14159265358979 * (fDia1 + fDia2) / 2.0
             + (fDia2 - fDia1) * (fDia2 - fDia1) / (4.0 * fCenter);   // L = 2C + π(D1+D2)/2 + ΔD²/(4C) / Pitch length
bValid := TRUE;                 // 有效回执 / Validity receipt
FC_DL_BeltLengthCalc := fBeltLength;   // 返回值 = 长度 / Return equals length
END_FUNCTION
